(* IEC 61131-3 sources: plcassist-cli/packages/volt-lsp-iec/test-corpus/pro2193/Device/Plc Logic/Application/09 Misc/Library Manager/L_MC2P_MotionControlCam, 92 files *)

(* ---- L_MC2P_CONSTANTS.gvl ---- *)
VAR_GLOBAL
	GC_DWCHECKIDCOND : DWORD := 1000;
	GC_DWCHECKIDCHAR : DWORD := 2000;
	GC_DWCHECKIDDATAXYA : DWORD := 3000;
	GC_DWCHECKIDDATAXY : DWORD := 3500;
	GC_DWCHECKIDDATAYA : DWORD := 4000;
	GC_DWCHECKIDDATAY : DWORD := 4500;
	GC_DWCHECKIDCAMDATA : DWORD := 5000;
	GC_DWCHECKIDSCCAMTABLEID : DWORD := 6000;
	GC_DWCHECKIDCAMID : DWORD := 7000;
	GC_DWCHECKIDCAMREF : DWORD := 12000;
	GC_DWCHECKIDTAPPET : DWORD := 8000;
	GC_DWCHECKIDTAPPETDATA : DWORD := 9000;
	GC_DWCHECKIDTAPPETREF : DWORD := 10000;
	GC_DWCHECKIDTAPPETID : DWORD := 11000;
	GC_DWCHECKIDTAPPETPOS : DWORD := 11001;
	GC_DWCHECKIDTAPPETTIME : DWORD := 11002;
	GC_LRCORRECTCONDITIONPOSITION : LREAL := 1E-06;
	GC_UIBLOCKEDNUMOFCYCLES : UINT := 10;
END_VAR

(* ---- L_MC2P_EVENTS.gvl ---- *)
VAR_GLOBAL
	CMPID_EVT_NEWCAMFILESDOWNLOADED : UDINT := 16#2003;
	EVT_CMPLENZEIPCSYSTEMNEWCAMFILESDOWNLOADED : UDINT := 16#10001;
	EVTPARAMID_CMPLENZEIPCSYSTEMNEWCAMFILESDOWNLOADED : UDINT := 16#1;
	EVTVERSION_CMPLENZEIPCSYSTEMNEWCAMFILESDOWNLOADED : UDINT := 16#1;
END_VAR

(* ---- L_MC2P_INTERNALCONST.gvl ---- *)
VAR_GLOBAL
	MAGICLML : DWORD := 16#46444D4C;
	MAGICCRPT : DWORD := 16#54505243;
	MAGICORGA : DWORD := 16#4147524F;
	MAGICEND : DWORD := 16#444E454C;
	MAGICCD : WORD := 16#4443;
	MAGICTD : WORD := 16#4454;
	C_CAM_CRC_BUFFERSIZE : DWORD := 96;
	CRC32TABLE : ARRAY [0..255] OF DWORD := [16#0, 16#77073096, 16#EE0E612C, 16#990951BA, 16#76DC419, 16#706AF48F, 16#E963A535, 16#9E6495A3, 16#EDB8832, 16#79DCB8A4, 16#E0D5E91E, 16#97D2D988, 16#9B64C2B, 16#7EB17CBD, 16#E7B82D07, 16#90BF1D91, 16#1DB71064, 16#6AB020F2, 16#F3B97148, 16#84BE41DE, 16#1ADAD47D, 16#6DDDE4EB, 16#F4D4B551, 16#83D385C7, 16#136C9856, 16#646BA8C0, 16#FD62F97A, 16#8A65C9EC, 16#14015C4F, 16#63066CD9, 16#FA0F3D63, 16#8D080DF5, 16#3B6E20C8, 16#4C69105E, 16#D56041E4, 16#A2677172, 16#3C03E4D1, 16#4B04D447, 16#D20D85FD, 16#A50AB56B, 16#35B5A8FA, 16#42B2986C, 16#DBBBC9D6, 16#ACBCF940, 16#32D86CE3, 16#45DF5C75, 16#DCD60DCF, 16#ABD13D59, 16#26D930AC, 16#51DE003A, 16#C8D75180, 16#BFD06116, 16#21B4F4B5, 16#56B3C423, 16#CFBA9599, 16#B8BDA50F, 16#2802B89E, 16#5F058808, 16#C60CD9B2, 16#B10BE924, 16#2F6F7C87, 16#58684C11, 16#C1611DAB, 16#B6662D3D, 16#76DC4190, 16#1DB7106, 16#98D220BC, 16#EFD5102A, 16#71B18589, 16#6B6B51F, 16#9FBFE4A5, 16#E8B8D433, 16#7807C9A2, 16#F00F934, 16#9609A88E, 16#E10E9818, 16#7F6A0DBB, 16#86D3D2D, 16#91646C97, 16#E6635C01, 16#6B6B51F4, 16#1C6C6162, 16#856530D8, 16#F262004E, 16#6C0695ED, 16#1B01A57B, 16#8208F4C1, 16#F50FC457, 16#65B0D9C6, 16#12B7E950, 16#8BBEB8EA, 16#FCB9887C, 16#62DD1DDF, 16#15DA2D49, 16#8CD37CF3, 16#FBD44C65, 16#4DB26158, 16#3AB551CE, 16#A3BC0074, 16#D4BB30E2, 16#4ADFA541, 16#3DD895D7, 16#A4D1C46D, 16#D3D6F4FB, 16#4369E96A, 16#346ED9FC, 16#AD678846, 16#DA60B8D0, 16#44042D73, 16#33031DE5, 16#AA0A4C5F, 16#DD0D7CC9, 16#5005713C, 16#270241AA, 16#BE0B1010, 16#C90C2086, 16#5768B525, 16#206F85B3, 16#B966D409, 16#CE61E49F, 16#5EDEF90E, 16#29D9C998, 16#B0D09822, 16#C7D7A8B4, 16#59B33D17, 16#2EB40D81, 16#B7BD5C3B, 16#C0BA6CAD, 16#EDB88320, 16#9ABFB3B6, 16#3B6E20C, 16#74B1D29A, 16#EAD54739, 16#9DD277AF, 16#4DB2615, 16#73DC1683, 16#E3630B12, 16#94643B84, 16#D6D6A3E, 16#7A6A5AA8, 16#E40ECF0B, 16#9309FF9D, 16#A00AE27, 16#7D079EB1, 16#F00F9344, 16#8708A3D2, 16#1E01F268, 16#6906C2FE, 16#F762575D, 16#806567CB, 16#196C3671, 16#6E6B06E7, 16#FED41B76, 16#89D32BE0, 16#10DA7A5A, 16#67DD4ACC, 16#F9B9DF6F, 16#8EBEEFF9, 16#17B7BE43, 16#60B08ED5, 16#D6D6A3E8, 16#A1D1937E, 16#38D8C2C4, 16#4FDFF252, 16#D1BB67F1, 16#A6BC5767, 16#3FB506DD, 16#48B2364B, 16#D80D2BDA, 16#AF0A1B4C, 16#36034AF6, 16#41047A60, 16#DF60EFC3, 16#A867DF55, 16#316E8EEF, 16#4669BE79, 16#CB61B38C, 16#BC66831A, 16#256FD2A0, 16#5268E236, 16#CC0C7795, 16#BB0B4703, 16#220216B9, 16#5505262F, 16#C5BA3BBE, 16#B2BD0B28, 16#2BB45A92, 16#5CB36A04, 16#C2D7FFA7, 16#B5D0CF31, 16#2CD99E8B, 16#5BDEAE1D, 16#9B64C2B0, 16#EC63F226, 16#756AA39C, 16#26D930A, 16#9C0906A9, 16#EB0E363F, 16#72076785, 16#5005713, 16#95BF4A82, 16#E2B87A14, 16#7BB12BAE, 16#CB61B38, 16#92D28E9B, 16#E5D5BE0D, 16#7CDCEFB7, 16#BDBDF21, 16#86D3D2D4, 16#F1D4E242, 16#68DDB3F8, 16#1FDA836E, 16#81BE16CD, 16#F6B9265B, 16#6FB077E1, 16#18B74777, 16#88085AE6, 16#FF0F6A70, 16#66063BCA, 16#11010B5C, 16#8F659EFF, 16#F862AE69, 16#616BFFD3, 16#166CCF45, 16#A00AE278, 16#D70DD2EE, 16#4E048354, 16#3903B3C2, 16#A7672661, 16#D06016F7, 16#4969474D, 16#3E6E77DB, 16#AED16A4A, 16#D9D65ADC, 16#40DF0B66, 16#37D83BF0, 16#A9BCAE53, 16#DEBB9EC5, 16#47B2CF7F, 16#30B5FFE9, 16#BDBDF21C, 16#CABAC28A, 16#53B39330, 16#24B4A3A6, 16#BAD03605, 16#CDD70693, 16#54DE5729, 16#23D967BF, 16#B3667A2E, 16#C4614AB8, 16#5D681B02, 16#2A6F2B94, 16#B40BBE37, 16#C30C8EA1, 16#5A05DF1B, 16#2D02EF8D];
	C_TAPPETS_BUFFERSIZE : DWORD := 23;
END_VAR

(* ---- L_MC2P_IMOTIONDATA.itf ---- *)
INTERFACE L_MC2P_IMOTIONDATA
END_INTERFACE

(* ---- L_MC2P_ITAPPETDATA.itf ---- *)
INTERFACE L_MC2P_ITAPPETDATA
END_INTERFACE

(* ---- L_MC2P_SETVALUES.itf ---- *)
INTERFACE L_MC2P_SETVALUES
END_INTERFACE

METHOD GETVALUES : LREAL
VAR_INPUT
	ESOURCE : MC_Source;
END_VAR
END_METHOD

(* ---- L_MC2P_TAPPET_REF.itf ---- *)
INTERFACE L_MC2P_TAPPET_REF
END_INTERFACE

METHOD GETID : DWORD
END_METHOD

METHOD GETTAPPETDATA : POINTER TO L_MC2P_TappetData
END_METHOD

METHOD SETCAMDATAACTIVE
VAR_INPUT
	XCAMACITVE : BOOL;
END_VAR
END_METHOD

METHOD SETMASTERVALUES
VAR_INPUT
	LRMASTERPOS : LREAL;
END_VAR
END_METHOD

(* ---- MC_CAM_REF.itf ---- *)
INTERFACE MC_CAM_REF
END_INTERFACE

METHOD GETCAMDATA : POINTER TO L_MC2P_CamData
END_METHOD

METHOD GETID : DWORD
END_METHOD

METHOD SETCAMDATAACTIVE
VAR_INPUT
	XCAMACITVE : BOOL;
END_VAR
END_METHOD

METHOD SETMASTERVALUES
VAR_INPUT
	LRMASTERPOS : LREAL;
END_VAR
END_METHOD

(* ---- GETBOOLEANPROPERTY.fun ---- *)
FUNCTION GETBOOLEANPROPERTY : BOOL
VAR_INPUT
	STKEY : WSTRING;
END_VAR
END_FUNCTION

(* ---- GETCOMPANY.fun ---- *)
FUNCTION GETCOMPANY : WSTRING
END_FUNCTION

(* ---- GETNUMBERPROPERTY.fun ---- *)
FUNCTION GETNUMBERPROPERTY : DINT
VAR_INPUT
	STKEY : WSTRING;
END_VAR
END_FUNCTION

(* ---- GETTEXTPROPERTY.fun ---- *)
FUNCTION GETTEXTPROPERTY : WSTRING
VAR_INPUT
	STKEY : WSTRING;
END_VAR
END_FUNCTION

(* ---- GETTEXTPROPERTY2.fun ---- *)
FUNCTION GETTEXTPROPERTY2 : POINTER TO WSTRING
VAR_INPUT
	STKEY : WSTRING;
END_VAR
END_FUNCTION

(* ---- GETTITLE.fun ---- *)
FUNCTION GETTITLE : WSTRING
END_FUNCTION

(* ---- GETVERSION.fun ---- *)
FUNCTION GETVERSION : VERSION
END_FUNCTION

(* ---- GETVERSIONPROPERTY.fun ---- *)
FUNCTION GETVERSIONPROPERTY : VERSION
VAR_INPUT
	STKEY : WSTRING;
END_VAR
END_FUNCTION

(* ---- L_MC2P_CAMGETDATA.fun ---- *)
FUNCTION L_MC2P_CAMGETDATA : POINTER TO BYTE
VAR_INPUT
	ITFCAMDATA : L_MC2P_IMotionData;
	IDX : UDINT;
	ECAMTYPE : L_MC2P_CamType;
END_VAR
END_FUNCTION

(* ---- L_MC2P_CAMGETDATA2.fun ---- *)
FUNCTION L_MC2P_CAMGETDATA2 : BOOL
VAR_INPUT
	ITFCAMDATA : L_MC2P_IMotionData;
	IDX1 : UDINT;
	IDX2 : UDINT;
	ECAMTYPE : L_MC2P_CamType;
END_VAR
VAR_OUTPUT
	PSCDATA1 : POINTER TO BYTE;
	PSCDATA2 : POINTER TO BYTE;
END_VAR
END_FUNCTION

(* ---- L_MC2P_CAMGETXVALUE2.fun ---- *)
FUNCTION L_MC2P_CAMGETXVALUE2 : BOOL
VAR_INPUT
	ITFCAMDATA : L_MC2P_IMotionData;
	IDX1 : UDINT;
	IDX2 : UDINT;
	ECAMTYPE : L_MC2P_CamType;
	LRMASTEP : LREAL;
	LRXSTART : LREAL;
END_VAR
VAR_OUTPUT
	LRX1 : LREAL;
	LRX2 : LREAL;
END_VAR
END_FUNCTION

(* ---- L_MC2P_CAMGETYVALUE2.fun ---- *)
FUNCTION L_MC2P_CAMGETYVALUE2 : BOOL
VAR_INPUT
	ITFCAMDATA : L_MC2P_IMotionData;
	IDX1 : UDINT;
	IDX2 : UDINT;
	ECAMTYPE : L_MC2P_CamType;
END_VAR
VAR_OUTPUT
	LRY1 : LREAL;
	LRY2 : LREAL;
END_VAR
END_FUNCTION

(* ---- L_MC2P_CHECK_CAMREFEQ.fun ---- *)
FUNCTION L_MC2P_CHECK_CAMREFEQ : BOOL
VAR_INPUT
	CAMREFNEW : MC_CAM_REF;
	CAMREFOLD : MC_CAM_REF;
END_VAR
END_FUNCTION

(* ---- L_MC2P_CHECK_CAMTABLECHANGED.fun ---- *)
FUNCTION L_MC2P_CHECK_CAMTABLECHANGED : BOOL
VAR_INPUT
	SCCAMTABLENEW : MC_Cam_REF;
	SCCAMTABLEOLD : MC_Cam_REF;
	SCCAMINFOOLD : L_MC2P_CamInfo;
END_VAR
END_FUNCTION

(* ---- L_MC2P_CHECK_CAMTABLEVALID.fun ---- *)
FUNCTION L_MC2P_CHECK_CAMTABLEVALID : BOOL
VAR_INPUT
	CAMTABLE : MC_Cam_REF;
END_VAR
END_FUNCTION

(* ---- L_MC2P_CONVERTPOSTOMODULOPOS.fun ---- *)
FUNCTION L_MC2P_CONVERTPOSTOMODULOPOS : LREAL
VAR_INPUT
	LRPOS : LREAL;
	LRPERIOD : LREAL;
END_VAR
END_FUNCTION

(* ---- L_MC2P_CONVERTPOSTOMODULOPOSEXTENDED.fun ---- *)
FUNCTION L_MC2P_CONVERTPOSTOMODULOPOSEXTENDED : LREAL
VAR_INPUT
	LRPOS : LREAL;
	LRPERIOD : LREAL;
END_VAR
END_FUNCTION

(* ---- L_MC2P_HLPMODULO.fun ---- *)
FUNCTION L_MC2P_HLPMODULO : LREAL
VAR_INPUT
	LRINPUT : LREAL;
	LRLENGHT : LREAL;
END_VAR
END_FUNCTION

(* ---- L_MC2P_HLPMODULOADD.fun ---- *)
FUNCTION L_MC2P_HLPMODULOADD : LREAL
VAR_INPUT
	LRINPUT : LREAL;
	LROFFSET : LREAL;
	LRLENGHT : LREAL;
END_VAR
END_FUNCTION

(* ---- L_MC2P_HLPMODULODIFF.fun ---- *)
FUNCTION L_MC2P_HLPMODULODIFF : LREAL
VAR_INPUT
	LRDIFF : LREAL;
	LRLEN : LREAL;
END_VAR
END_FUNCTION

(* ---- L_MC2P_HLPMODULOZERO.fun ---- *)
FUNCTION L_MC2P_HLPMODULOZERO : BOOL
VAR_INPUT
	LRDIFF : LREAL;
	LRLEN : LREAL;
END_VAR
END_FUNCTION

(* ---- CRYPTING.fb ---- *)
FUNCTION_BLOCK CRYPTING
END_FUNCTION_BLOCK

METHOD DECRYPTMODE1
VAR_INPUT
	NUM_CYCLES : WORD;
	V : POINTER TO ARRAY [0..1] OF UDINT;
	K : ARRAY [0..3] OF UDINT;
END_VAR
END_METHOD

METHOD DECRYPTMODE64
VAR_INPUT
	NUM_CYCLES : WORD;
	V : POINTER TO ARRAY [0..1] OF ULINT;
	K : ARRAY [0..3] OF ULINT;
END_VAR
END_METHOD

METHOD ENCRYPTMODE1
VAR_INPUT
	NUM_CYCLES : WORD;
	V : POINTER TO ARRAY [0..1] OF UDINT;
	K : ARRAY [0..3] OF UDINT;
END_VAR
END_METHOD

METHOD ENCRYPTMODE64
VAR_INPUT
	NUM_CYCLES : WORD;
	V : POINTER TO ARRAY [0..1] OF ULINT;
	K : ARRAY [0..3] OF ULINT;
END_VAR
END_METHOD

METHOD GETLINTFROMCHAR : ULINT
VAR_INPUT
	ABDATA : ARRAY [0..3] OF BYTE;
END_VAR
END_METHOD

METHOD SETKEY : ARRAY [0..3] OF ULINT
VAR_INPUT
	SSTRING : STRING(16);
END_VAR
END_METHOD

(* ---- GLOBALTEXTLIST.fb ---- *)
FUNCTION_BLOCK GLOBALTEXTLIST
VAR
	M_TEXTLISTFILE : STRING(255);
	_STNAMESPACE : STRING;
END_VAR
END_FUNCTION_BLOCK

(* ---- IMAGEPOOL.fb ---- *)
FUNCTION_BLOCK IMAGEPOOL
VAR
	M_STNAMESPACE : STRING(80);
	M_STHELPVARID : STRING;
	M_STHELPVARPATH : STRING(255);
	M_STHELP : STRING;
	M_REGISTERIMAGES : BOOL := TRUE;
END_VAR
END_FUNCTION_BLOCK

METHOD FB_INIT : BOOL
VAR_INPUT
	BINITRETAINS : BOOL;
	BINCOPYCODE : BOOL;
END_VAR
END_METHOD

METHOD FB_REINIT : BOOL
END_METHOD

METHOD FB_EXIT : BOOL
VAR_INPUT
	BINCOPYCODE : BOOL;
END_VAR
END_METHOD

(* ---- L_MC2P_AXISCONVERTERBASE.fb ---- *)
FUNCTION_BLOCK L_MC2P_AXISCONVERTERBASE EXTENDS L_MC2P_CamAxisConverter
VAR_INPUT
	XENABLE : BOOL;
	LRCYCMASTERPOS : LREAL;
	LRCYCMASTERVEL : LREAL;
	LRCYCMASTERACC : LREAL;
	LRCYCLELENGTHMASTER : LREAL := 360;
	IMASTERMOVEMENTTYPE : INT := 0;
	LRCYCLELENGTHSLAVE : LREAL := 360;
	ISLAVEMOVEMENTTYPE : INT := 0;
	LRSETOFFSET : LREAL;
	LRSETSCALING : LREAL := 1;
	ESCALINGMODE : L_MC2P_ScalingMode := L_MC2P_ScalingMode.absolute;
END_VAR
VAR_OUTPUT
	XERROR : BOOL;
	EERRORID : L_IE1P_Error;
	XBUSY : BOOL;
	LRSETSLAVEPOSOUT : LREAL;
	LRSETSLAVEVELOUT : LREAL;
	LRSETSLAVEACCOUT : LREAL;
END_VAR
VAR
	XERROR_OLD : BOOL;
	EERRORID_OLD : L_IE1P_Error;
	XENABLE_OLD : BOOL;
	LRCYCMASTERPOS_OLD : LREAL;
	ESTATE : L_MC2P_States := L_MC2P_States.INIT;
	XSTATEENTRY : BOOL;
	BYCONVERTERMODE : BYTE;
	SCSETSLAVEOUT : L_MC2P_AxisProfile;
END_VAR
END_FUNCTION_BLOCK

METHOD CALL_CONVERTLINEARTOLINEAR
END_METHOD

METHOD CALL_CONVERTLINEARTOMODULO
END_METHOD

METHOD CALL_CONVERTMODULOTOLINEAR
END_METHOD

METHOD CALL_CONVERTMODULOTOMODULO
END_METHOD

METHOD CALL_ERRORHANDLER
END_METHOD

METHOD CALL_FBMETHODS
END_METHOD

METHOD CALL_OUTPUT
END_METHOD

METHOD CALL_RESETCOMMANDS
END_METHOD

METHOD CALL_RESETOUTPUT
END_METHOD

METHOD CALL_STATEMASHINE
END_METHOD

METHOD CALL_S000_CYCLIC
END_METHOD

METHOD CALL_S001_INIT
END_METHOD

METHOD CALL_S010_READY
END_METHOD

METHOD CALL_S200_SYNCHRON
END_METHOD

METHOD CALL_S998_ERROR
END_METHOD

(* ---- L_MC2P_BOUNDSCAM.fb ---- *)
FUNCTION_BLOCK L_MC2P_BOUNDSCAM EXTENDS L_MC2P_TemplateSlaveAxis
VAR_INPUT
	XEXECUTE : BOOL;
	ITFCAMTABLE : MC_CAM_REF;
	LRMAVEL : LREAL;
	LRMAACC : LREAL;
	UDINUMOFPOINTS : UDINT;
	UDIPOINTSPERCYCLE : UDINT;
END_VAR
VAR_OUTPUT
	XDONE : BOOL;
	XBUSY : BOOL;
	XERROR : BOOL;
	EERRORID : L_IE1P_Error;
	LRPOSMAX : LREAL;
	LRPOSMIN : LREAL;
	LRVELMAX : LREAL;
	LRVELMIN : LREAL;
	LRACCDECMAX : LREAL;
	LRACCDECMIN : LREAL;
END_VAR
VAR
	L_MC2P_CAMBASIC1 : L_MC2P_CamBasic;
	SCVIRTUALSLAVE : L_MC2P_AxisProfile;
	I : UDINT;
	LRMASTEP : LREAL;
	LRMAPOS : LREAL;
	XBREAK : BOOL;
	XEXECUTEOLD : BOOL;
	XRESETOUTPUT : BOOL;
	SCVIRTUALMASTER : L_MC2P_AxisProfile;
	LRMAVEL_INT : LREAL;
	LRMAACC_INT : LREAL;
	UDINUMOFPOINTS_INT : UDINT := 2;
	UDIPOINTSPERCYCLE_INT : UDINT;
	PCAMDATA_INT : POINTER TO L_MC2P_CamData;
	SCCAMINFO : L_MC2P_CamInfo;
	LRPOSMAX_INT : LREAL;
	LRPOSMIN_INT : LREAL;
	LRVELMAX_INT : LREAL;
	LRVELMIN_INT : LREAL;
	LRACCDECMAX_INT : LREAL;
	LRACCDECMIN_INT : LREAL;
END_VAR
END_FUNCTION_BLOCK

METHOD READINPUTS
END_METHOD

METHOD RESET_MINMAXVALUES
END_METHOD

METHOD RESET_OUTPUTS
END_METHOD

METHOD RESET_OUTPUTSBYERROR
END_METHOD

METHOD SET_MINMAXVALUES
END_METHOD

(* ---- L_MC2P_CAMAXISCONVERTER.fb ---- *)
FUNCTION_BLOCK L_MC2P_CAMAXISCONVERTER
VAR
	_XERROR : BOOL;
	LRSLAVEPERIOD_INT : LREAL := 0;
	LRSETSLAVEPOSOUTSCALED : LREAL := 0;
	DWACTSLAVEPOS_INT : DWORD := 0;
	LRSETSLAVEPOSOUT_INT : LREAL := 0;
	LRSLAVEOFFSET_INT : LREAL := 0;
	LRSLAVEOFFSET_REL : LREAL := 0;
	LRYOFFSET_INT : LREAL := 0;
	LRSETYPOS_INT : LREAL := 0;
	LRSETYPOS_SCALED : LREAL := 0;
	LRSETYSCALING_INT : LREAL := 1;
	ALRMEM : ARRAY [1..7] OF LREAL;
	XMODULOMODE : BOOL;
	LRXPERIOD_NEXT : LREAL;
	LRSTARTXAXIS_NEXT : LREAL := 0;
	LRSETXPOSOUT_MODULO : LREAL := 0;
	LRSETXPOSOUT_MODULO_OLD : LREAL := 0;
	LRSETXPOSOUT_INT : LREAL := 0;
	LRXPERIOD_INT : LREAL := 0;
	LRSTARTXAXIS_INT : LREAL := 0;
	LRSETXSCALING_INT : LREAL := 1;
	LROFFSET_INT : LREAL := 0;
	LROFFSET_REL : LREAL := 0;
	LRONECYCLEXOFFSET_INT : LREAL := 0;
	XLOADSTARTXPOS : BOOL;
	LRLOADSTARTXPOS : LREAL;
	XCHECKMASTERPOSBYLOAD : BOOL;
	LRCYCSETMASTERPOSBYLOAD : LREAL;
	LRSETXPOSBYLOAD : LREAL;
	XOVERRUNMASTERPOS : BOOL := FALSE;
	XOVERRUNMASTERNEG : BOOL := FALSE;
	LWREMAINDER_ADD : LWORD := 0;
	LWREMAINDER_INT : LWORD := 0;
	LRREMAINDER_INT : LREAL := 0;
	LRCYCSETMASTERPOS_VIRTUAL : LREAL := 0;
	LRMASTERPERIOD_VIRTUAL : LREAL := 0;
	IPERIODFACTOR : INT := 0;
	IPERIODCTN : INT := 0;
	LRCYCSETMASTERVEL_INT : LREAL;
	LRCYCSETMASTERPOS_INT : LREAL;
	LRMASTERPERIOD_INT : LREAL := 0;
	LRCYCSETMASTERPOS_SCALED : LREAL := 0;
	LRMASTERPERIOD_SCALED : LREAL := 0;
	XEOP_INIT : BOOL := TRUE;
	IEOP_CYCLECNTR : INT := 0;
	IEOP_CYCLECNTR2 : INT := 0;
	LWEOP_TCHECKSUM : LWORD;
	XEOP_ENDOFPERIODPOSITIVE : BOOL;
	XEOP_ENDOFPERIODNEGATIVE : BOOL;
	WEOP_STEPPER : WORD := 0;
	LREOP_CYCSETMASTERPOS_OLD : LREAL;
	LREOP_SETXPOSOUT_MODULO_OLD : LREAL;
	LREOP_XPERIOD : LREAL;
	LREOP_XPERIOD_OLD : LREAL;
	XEOP_ENDOFPROFPOSITIVE : BOOL;
	XEOP_ENDOFPROFNEGATIVE : BOOL;
	LREOP_SETXDELTAPOS : LREAL;
	LREOP_SETXDELTA2POS : LREAL;
	LREOP_SETXDELTA3POS : LREAL;
	LREOP_SETXDELTAPOS_OLD : LREAL;
	LREOP_SETXDELTA2POS_OLD : LREAL;
	LREOP_SETXSCALING_OLD : LREAL;
	LREOP_OFFSET_OLD : LREAL;
	ALREOP_MEM : ARRAY [1..7] OF LREAL;
	XEOP_RAMPOFFSETMODE : BOOL;
	XEOP_RAMPSCALINGMODE : BOOL;
	XOUTOFCAMPOSITIVE_INT : BOOL;
	XOUTOFCAMNEGATIVE_INT : BOOL;
	LRTEMP : LREAL;
	LRENDOFPROFILEFACTOR_INT : LREAL := 1;
	LRCYCSETMASTERPOSATSCLING0 : LREAL;
	LRSETXPOSOUTATSCLING0 : LREAL;
	LRSETXSCALINGATSCLING0 : LREAL;
	LRDWUPPERLIMIT : LREAL := 16#FFFFFFFF;
	DWDWUPPERLIMIT : DWORD := 16#FFFFFFFF;
	LRLWUPPERLIMIT : LREAL := 16#7FFFFFFFFFFFFFFF;
	LWENDOFPROFILECHECKSUM : LWORD;
END_VAR
END_FUNCTION_BLOCK

METHOD CALC_LRSETSLAVEPOSOUT : LREAL
VAR_IN_OUT
	LRSETYPOS : LREAL;
END_VAR
END_METHOD

METHOD CALC_LRSETXLINPOSOUT : LREAL
VAR_IN_OUT
	LRCYCSETMASTERPOS : LREAL;
	LRCYCSETMASTERVEL : LREAL;
	LRCYCSETMASTERACC : LREAL;
END_VAR
END_METHOD

METHOD CALC_LRSETXPOSOUT : LREAL
VAR_IN_OUT
	LRCYCSETMASTERPOS : LREAL;
	LRCYCSETMASTERVEL : LREAL;
	LRCYCSETMASTERACC : LREAL;
END_VAR
END_METHOD

METHOD CALC_LRSETXPOSOUTEXTENDED : LREAL
VAR_INPUT
	LRENDOFPROFILEWINDOW : LREAL;
END_VAR
VAR_OUTPUT
	LRSETXPOSOUT : LREAL;
	XENDOFPROFPOSITIVE : BOOL;
	XENDOFPROFNEGATIVE : BOOL;
	XEXTRAPOLATECAM : BOOL;
	XCYCLEZERO : BOOL;
	XOUTOFCAMPOSITIVE : BOOL;
	XOUTOFCAMNEGATIVE : BOOL;
END_VAR
VAR_IN_OUT
	LRCYCSETMASTERPOS : LREAL;
	LRCYCSETMASTERPOS_OLD : LREAL;
	LRCYCSETMASTERVEL : LREAL;
	LRCYCSETMASTERACC : LREAL;
END_VAR
END_METHOD

METHOD CALL_RESET
END_METHOD

METHOD SET_LRENDOFPROFILEFACTOR : BOOL
VAR_INPUT
	LRIN : LREAL;
END_VAR
END_METHOD

METHOD CALC_DWADDMODULO : DWORD
VAR_INPUT
	LRSETXPOS : LREAL;
	LRSETYPOS : LREAL;
	LRPERIOD : LREAL;
END_VAR
END_METHOD

METHOD CALC_DWSUBMODULO : DWORD
VAR_INPUT
	LRSETYPOS : LREAL;
	LRSETXPOS : LREAL;
	LRPERIOD : LREAL;
END_VAR
END_METHOD

METHOD CALC_LRADDMODULO : LREAL
VAR_INPUT
	LRSETXPOS : LREAL;
	LRSETYPOS : LREAL;
	LRPERIOD : LREAL;
END_VAR
END_METHOD

METHOD CALC_LRSUBMODULO : LREAL
VAR_INPUT
	LRSETXPOS : LREAL;
	LRSETYPOS : LREAL;
	LRPERIOD : LREAL;
END_VAR
END_METHOD

METHOD CALL_CHECKLOADXPOSAFTERCONVERTER
END_METHOD

METHOD CALL_CHECKMODULOOVERRUN
VAR_IN_OUT
	LRSETPOS : LREAL;
	LRSETVEL : LREAL;
	LRPERIOD : LREAL;
	XOVERRUNPOS : BOOL;
	XOVERRUNNEG : BOOL;
	ALRMEM : ARRAY [1..7] OF LREAL;
END_VAR
END_METHOD

METHOD CALL_DWCONVERTLREALTODWORD : DWORD
VAR_INPUT
	LRIN : LREAL;
	LRPERIOD : LREAL;
END_VAR
END_METHOD

METHOD CALL_DWCONVERTLREALTOLWORD : LWORD
VAR_INPUT
	LRIN : LREAL;
	LRPERIOD : LREAL;
END_VAR
END_METHOD

METHOD CALL_LRCONVERTDWORDTOLREAL : LREAL
VAR_INPUT
	DWIN : DWORD;
	LRPERIOD : LREAL;
END_VAR
END_METHOD

METHOD CALL_LRCONVERTLREALTOMODULO : LREAL
VAR_INPUT
	LRIN : LREAL;
	LRPERIOD : LREAL;
END_VAR
END_METHOD

METHOD CALL_LRCONVERTLWORDTOLREAL : LREAL
VAR_INPUT
	LWIN : LWORD;
	LRPERIOD : LREAL;
END_VAR
END_METHOD

METHOD CALC_MASTERVIRTUALPERIOD
END_METHOD

METHOD CALL_CHECKMODULOMODE
END_METHOD

METHOD CALL_CHECKZERROPOS
VAR_INPUT
	LRCYCSETMASTERPOS : LREAL;
END_VAR
END_METHOD

METHOD CHECK_XENDOFPROFILE : BOOL
VAR_INPUT
	LRSETXPOS : LREAL;
	LRSETXDELTAPOS : LREAL;
	LRSETXDELTA2POS : LREAL;
	LRSETXDELTA3POS : LREAL;
	LRXSTART : LREAL;
	LRXEND : LREAL;
	LRXPERIOD : LREAL;
END_VAR
VAR_OUTPUT
	LRSETNEXTXPOSOUT : LREAL;
	XPOSITIVE : BOOL;
	XNEGATIVE : BOOL;
END_VAR
END_METHOD

METHOD CALL_XMASTERVALID : BOOL
END_METHOD

METHOD GET_LRSLAVEOFFSETREL : LREAL
END_METHOD

METHOD GET_LRXOFFSETREL : LREAL
END_METHOD

METHOD LOAD_STARTXPOS
VAR_IN_OUT
	LRLOADXPOS : LREAL;
	LRCYCSETMASTERPOS : LREAL;
END_VAR
END_METHOD

METHOD SET_ACTAXISLIMIT
VAR_IN_OUT
	LRSTARTXAXIS : LREAL := 0;
	LRENDXAXIS : LREAL := 0;
END_VAR
END_METHOD

METHOD SET_EOPXOFFSETMODE
VAR_INPUT
	XRAMPOFFSETMODE : BOOL;
END_VAR
END_METHOD

METHOD SET_EOPXSCALINGMODE
VAR_INPUT
	XRAMPSCALINGMODE : BOOL;
END_VAR
END_METHOD

METHOD SET_NEWXPERIOD
VAR_IN_OUT
	LRSETXPOSOUT : LREAL;
	LRSETXPERIOD : LREAL;
	LRCYCSETMASTERPOS : LREAL;
END_VAR
END_METHOD

METHOD SET_NEXTAXISLIMIT
VAR_IN_OUT
	LRSTARTXAXIS : LREAL := 0;
	LRENDXAXIS : LREAL := 0;
END_VAR
END_METHOD

METHOD SET_ONECYCLEOFFSET
VAR_INPUT
	LRXOFFSET : LREAL;
END_VAR
END_METHOD

METHOD SET_XAXISLIMIT
VAR_INPUT
	LRSTARTXAXIS : LREAL;
	LRENDXAXIS : LREAL;
	LRSETSCALING : LREAL;
END_VAR
END_METHOD

METHOD SET_XOFFSET
VAR_INPUT
	LRSETOFFSET : LREAL;
END_VAR
END_METHOD

METHOD SET_XPERIOD
VAR_IN_OUT
	LRXPERIOD : LREAL;
	LRSETSCALING : LREAL;
END_VAR
END_METHOD

METHOD SET_XPOSTOMASTERPOS : DWORD
VAR_IN_OUT
	LRCYCSETMASTERPOS : LREAL;
END_VAR
END_METHOD

METHOD SET_XSCALING
VAR_INPUT
	LRSETSCALING : LREAL := 1;
	WSCALINGMODE : WORD := 0;
	LRCYCSETMASTERPOS : LREAL;
	LRCYCSETMASTERPOS_OLD : LREAL;
END_VAR
END_METHOD

METHOD SET_LRMASTERPERIOD
VAR_INPUT
	LRSETMASTERPERIOD : LREAL;
END_VAR
END_METHOD

METHOD LOAD_SALVEPOS
VAR_INPUT
	LRLOADSLAVEPOS : LREAL;
	LRSETYPOS : LREAL;
	LRSETYSCALING : LREAL;
END_VAR
END_METHOD

METHOD SET_SLAVEPOSTOYPOS : DWORD
VAR_INPUT
	LRSETYSCALING : LREAL;
END_VAR
END_METHOD

METHOD SET_YSCALING
VAR_INPUT
	LRSETSCALING : LREAL := 1;
	WSCALINGMODE : WORD := 0;
	LRSETSLAVEPOSOUT : LREAL;
	LRSETYPOS_OLD : LREAL;
END_VAR
END_METHOD

METHOD SET_LRCAMPOSDIFF
VAR_INPUT
	LRCAMPOSDIFF : LREAL;
END_VAR
END_METHOD

METHOD SET_LRCAMSWITCHREL
VAR_INPUT
	XDIRECTIONPOS : BOOL;
	LRYSCALINGEND : LREAL;
	LRYSCALINGSTART : LREAL;
	LRCAMYEND : LREAL;
	LRCAMYSTART : LREAL;
END_VAR
END_METHOD

METHOD SET_LRSLAVEOFFSET
VAR_INPUT
	LRSETOFFSET : LREAL;
END_VAR
END_METHOD

METHOD SET_LRSLAVEPERIOD
VAR_INPUT
	LRSETSLAVEPERIOD : LREAL;
END_VAR
END_METHOD

METHOD SET_LRYOFFSET
VAR_INPUT
	LRSETOFFSET : LREAL;
END_VAR
END_METHOD

(* ---- L_MC2P_CAMBASIC.fb ---- *)
FUNCTION_BLOCK L_MC2P_CAMBASIC
VAR
	LRENDVEL : LREAL;
	LRSTARTVEL : LREAL;
	LRENDACC : LREAL;
	LRSTARTACC : LREAL;
	LRMASTEP : LREAL;
	UDISEG : UDINT;
	UDISEGOLD : UDINT;
	UDISEGADD2 : UDINT;
	UDISEGSUB1 : UDINT;
	UDILEFTBORDER : UDINT;
	UDIRIGHTBORDER : UDINT;
	XFOUNDSEG : BOOL;
	SCCHAR : ARRAY [0..1] OF L_MC2P_Characteristics;
	WDEBUG : WORD;
	XRESTARTSERCH : BOOL;
	LRMAPOSOLD : LREAL;
	PCAMDATAOLD : POINTER TO BYTE;
	PDATAOLD : POINTER TO BYTE;
	ECAMTYPEOLD : DWORD;
	UDINUMOFELEMENTSOLD : DWORD;
	LRXSTARTPOSOLD : LREAL;
	LRXENDPOSOLD : LREAL;
	WSLAVESTATEOLDCYCLE : WORD;
	WSLAVESTATEOLDCAM : WORD;
	SCOUTPUTSLAVEOLDCYCLE : L_MC2P_AxisProfile;
	XNEWCAMDETECTED : BOOL;
	ACTUALSEGMENT : UDINT;
	FOUNDSEG : BOOL;
END_VAR
END_FUNCTION_BLOCK

METHOD CALCULATECAMPROFILE
VAR_INPUT
	PCAMDATA : POINTER TO L_MC2P_CamData;
	SCINPUTMASTER : L_MC2P_AxisProfile;
	XPERIODIC : BOOL;
	XEXTRAPOLATECAM : BOOL;
END_VAR
VAR_OUTPUT
	SCOUTPUTSLAVE : L_MC2P_AxisProfile;
	XERROR : BOOL;
	EERRORID : L_IE1P_Error;
END_VAR
END_METHOD

METHOD CALCULATECAMPROFILEINT
VAR_INPUT
	PCAMDATA : POINTER TO L_MC2P_CamData;
	SCINPUTMASTER : L_MC2P_AxisProfile;
	XPERIODIC : BOOL;
END_VAR
VAR_OUTPUT
	SCOUTPUTSLAVE : L_MC2P_AxisProfile;
	XERROR : BOOL;
	EERRORID : L_IE1P_Error;
END_VAR
END_METHOD

METHOD CAMGENERATORCOND
VAR_INPUT
	ITFCAMDATA : L_MC2P_IMotionData;
	LRINPUTMASTERVEL : LREAL;
	PSCCHAR : POINTER TO L_MC2P_Characteristics;
END_VAR
VAR_OUTPUT
	XERROR : BOOL;
	EERRORID : L_IE1P_Error;
END_VAR
END_METHOD

METHOD CAMPROFILERCHARCALC
VAR_INPUT
	PSCCHAR : POINTER TO L_MC2P_Characteristics;
	LRPOS : LREAL;
	UDISEGCHAR : UDINT;
	LRINPUTMASTERVEL : LREAL;
	LRINPUTMASTERACC : LREAL;
END_VAR
VAR_OUTPUT
	SCOUTPUTSLAVE : L_MC2P_AxisProfile;
END_VAR
END_METHOD

METHOD CAMPROFILERCHARSEARCH
VAR_INPUT
	PSCCHAR : POINTER TO L_MC2P_Characteristics;
	LRINPUTMASTERPOS : LREAL;
	ECAMTYPE : L_MC2P_CamType;
END_VAR
VAR_OUTPUT
	LRPOS : LREAL;
	UDISEGCHAR : UDINT;
END_VAR
END_METHOD

METHOD CAMPROFILERDATAEQUIY
VAR_INPUT
	PCAMDATA : POINTER TO L_MC2P_CamData;
	LRINPUTMASTERPOS : LREAL;
	LRINPUTMASTERVEL : LREAL;
	LRINPUTMASTERACC : LREAL;
	XPERIODIC : BOOL;
END_VAR
VAR_OUTPUT
	SCOUTPUTSLAVE : L_MC2P_AxisProfile;
	XERROR : BOOL;
	EERRORID : L_IE1P_Error;
END_VAR
END_METHOD

METHOD CAMPROFILERDATAEQUIYA
VAR_INPUT
	PCAMDATA : POINTER TO L_MC2P_CamData;
	LRINPUTMASTERPOS : LREAL;
	LRINPUTMASTERVEL : LREAL;
	LRINPUTMASTERACC : LREAL;
	XPERIODIC : BOOL;
END_VAR
VAR_OUTPUT
	SCOUTPUTSLAVE : L_MC2P_AxisProfile;
	XERROR : BOOL;
	EERRORID : L_IE1P_Error;
END_VAR
END_METHOD

METHOD CAMPROFILERDATANONEQUIXY
VAR_INPUT
	PCAMDATA : POINTER TO L_MC2P_CamData;
	LRINPUTMASTERPOS : LREAL;
	LRINPUTMASTERVEL : LREAL;
	LRINPUTMASTERACC : LREAL;
	XPERIODIC : BOOL;
END_VAR
VAR_OUTPUT
	SCOUTPUTSLAVE : L_MC2P_AxisProfile;
	XERROR : BOOL;
	EERRORID : L_IE1P_Error;
END_VAR
END_METHOD

METHOD CAMPROFILERDATANONEQUIXYA
VAR_INPUT
	PCAMDATA : POINTER TO L_MC2P_CamData;
	LRINPUTMASTERPOS : LREAL;
	LRINPUTMASTERVEL : LREAL;
	LRINPUTMASTERACC : LREAL;
	XPERIODIC : BOOL;
END_VAR
VAR_OUTPUT
	SCOUTPUTSLAVE : L_MC2P_AxisProfile;
	XERROR : BOOL;
	EERRORID : L_IE1P_Error;
END_VAR
END_METHOD

METHOD GETSTARTENDVALUES
VAR_INPUT
	PCAMDATA : POINTER TO L_MC2P_CamData;
END_VAR
VAR_OUTPUT
	LRSTARTSLAVE : LREAL;
	LRENDSLAVE : LREAL;
END_VAR
END_METHOD

METHOD RESETSEGMENT
END_METHOD

METHOD SEARCHSEGMENT
VAR_INPUT
	PCAMDATA : POINTER TO L_MC2P_CamData;
	LRINPUTMASTERPOS : LREAL;
	LRINPUTMASTERVEL : LREAL;
	XPERIODIC : BOOL;
END_VAR
VAR_OUTPUT
	XERROR : BOOL;
	EERRORID : L_IE1P_Error;
END_VAR
END_METHOD

METHOD FB_INIT : BOOL
VAR_INPUT
	BINITRETAINS : BOOL;
	BINCOPYCODE : BOOL;
END_VAR
END_METHOD

METHOD GETEXTREMVALUES_POLY5
VAR_INPUT
	PSCCHARCLUTCH : POINTER TO L_MC2P_Characteristics;
END_VAR
VAR_OUTPUT
	LRFSMAX1 : LREAL;
	LRFSMAX2 : LREAL;
	LRFSMAX3 : LREAL;
END_VAR
END_METHOD

METHOD GEN_BB_POLY5
VAR_INPUT
	PSCCONDLEFT : POINTER TO L_MC2P_XYVA;
	PSCCONDRIGHT : POINTER TO L_MC2P_XYVA;
	PSCCHAR : POINTER TO L_MC2P_Characteristics;
END_VAR
END_METHOD

METHOD GEN_BB_POLY7
VAR_INPUT
	PSCCONDLEFT : POINTER TO L_MC2P_XYVA;
	PSCCONDRIGHT : POINTER TO L_MC2P_XYVA;
	PSCCHAR : POINTER TO L_MC2P_Characteristics;
END_VAR
END_METHOD

METHOD GEN_GG_GERADE
VAR_INPUT
	PSCCONDLEFT : POINTER TO L_MC2P_XYVA;
	PSCCONDRIGHT : POINTER TO L_MC2P_XYVA;
	PSCCHAR : POINTER TO L_MC2P_Characteristics;
END_VAR
END_METHOD

METHOD GEN_GG_MODSIN
VAR_INPUT
	PSCCONDLEFT : POINTER TO L_MC2P_XYVA;
	PSCCONDRIGHT : POINTER TO L_MC2P_XYVA;
	PSCCHAR : POINTER TO L_MC2P_Characteristics;
END_VAR
END_METHOD

METHOD GEN_GG_POLY3
VAR_INPUT
	PSCCONDLEFT : POINTER TO L_MC2P_XYVA;
	PSCCONDRIGHT : POINTER TO L_MC2P_XYVA;
	PSCCHAR : POINTER TO L_MC2P_Characteristics;
END_VAR
END_METHOD

METHOD GEN_GR_POLY2
VAR_INPUT
	PSCCONDLEFT : POINTER TO L_MC2P_XYVA;
	PSCCONDRIGHT : POINTER TO L_MC2P_XYVA;
	PSCCHAR : POINTER TO L_MC2P_Characteristics;
END_VAR
END_METHOD

METHOD GEN_GU_HARMKOMB
VAR_INPUT
	PSCCONDLEFT : POINTER TO L_MC2P_XYVA;
	PSCCONDRIGHT : POINTER TO L_MC2P_XYVA;
	PSCCHAR : POINTER TO L_MC2P_Characteristics;
END_VAR
END_METHOD

METHOD GEN_RG_POLY2
VAR_INPUT
	PSCCONDLEFT : POINTER TO L_MC2P_XYVA;
	PSCCONDRIGHT : POINTER TO L_MC2P_XYVA;
	PSCCHAR : POINTER TO L_MC2P_Characteristics;
END_VAR
END_METHOD

METHOD GEN_RR_BESCHLTRAPEZ
VAR_INPUT
	PSCCONDLEFT : POINTER TO L_MC2P_XYVA;
	PSCCONDRIGHT : POINTER TO L_MC2P_XYVA;
	PSCCHAR : POINTER TO L_MC2P_Characteristics;
END_VAR
END_METHOD

METHOD GEN_RR_GENSIN
VAR_INPUT
	PSCCONDLEFT : POINTER TO L_MC2P_XYVA;
	PSCCONDRIGHT : POINTER TO L_MC2P_XYVA;
	PSCCHAR : POINTER TO L_MC2P_Characteristics;
END_VAR
END_METHOD

METHOD GEN_RR_MODBESCHLTRAPEZ
VAR_INPUT
	PSCCONDLEFT : POINTER TO L_MC2P_XYVA;
	PSCCONDRIGHT : POINTER TO L_MC2P_XYVA;
	PSCCHAR : POINTER TO L_MC2P_Characteristics;
END_VAR
END_METHOD

METHOD GEN_RR_QUADPARABEL
VAR_INPUT
	PSCCONDLEFT : POINTER TO L_MC2P_XYVA;
	PSCCONDRIGHT : POINTER TO L_MC2P_XYVA;
	PSCCHAR : POINTER TO L_MC2P_Characteristics;
END_VAR
END_METHOD

METHOD GEN_RR_SIN
VAR_INPUT
	PSCCONDLEFT : POINTER TO L_MC2P_XYVA;
	PSCCONDRIGHT : POINTER TO L_MC2P_XYVA;
	PSCCHAR : POINTER TO L_MC2P_Characteristics;
END_VAR
END_METHOD

METHOD GEN_RU_MODBESCHLTRAPEZ
VAR_INPUT
	PSCCONDLEFT : POINTER TO L_MC2P_XYVA;
	PSCCONDRIGHT : POINTER TO L_MC2P_XYVA;
	PSCCHAR : POINTER TO L_MC2P_Characteristics;
END_VAR
END_METHOD

METHOD GEN_UG_HARMKOMB
VAR_INPUT
	PSCCONDLEFT : POINTER TO L_MC2P_XYVA;
	PSCCONDRIGHT : POINTER TO L_MC2P_XYVA;
	PSCCHAR : POINTER TO L_MC2P_Characteristics;
END_VAR
END_METHOD

METHOD GEN_UR_MODBESCHLTRAPEZ
VAR_INPUT
	PSCCONDLEFT : POINTER TO L_MC2P_XYVA;
	PSCCONDRIGHT : POINTER TO L_MC2P_XYVA;
	PSCCHAR : POINTER TO L_MC2P_Characteristics;
END_VAR
END_METHOD

METHOD GEN_UU_SINGERKOMB : ARRAY [0..1] OF L_MC2P_Characteristics
VAR_INPUT
	PSCCONDLEFT : POINTER TO L_MC2P_XYVA;
	PSCCONDRIGHT : POINTER TO L_MC2P_XYVA;
	PSCCHAR : POINTER TO L_MC2P_Characteristics;
END_VAR
END_METHOD

METHOD PROF_BB_POLY5
VAR_INPUT
	PSCCHAR : POINTER TO L_MC2P_Characteristics;
	LRPOS : LREAL;
	PSCNORMSLAVE : POINTER TO L_MC2P_AxisProfile;
END_VAR
END_METHOD

METHOD PROF_BB_POLY7
VAR_INPUT
	PSCCHAR : POINTER TO L_MC2P_Characteristics;
	LRPOS : LREAL;
	PSCNORMSLAVE : POINTER TO L_MC2P_AxisProfile;
END_VAR
END_METHOD

METHOD PROF_GG_GERADE
VAR_INPUT
	PSCCHAR : POINTER TO L_MC2P_Characteristics;
	LRPOS : LREAL;
	PSCNORMSLAVE : POINTER TO L_MC2P_AxisProfile;
END_VAR
END_METHOD

METHOD PROF_GG_MODSIN
VAR_INPUT
	PSCCHAR : POINTER TO L_MC2P_Characteristics;
	LRPOS : LREAL;
	PSCNORMSLAVE : POINTER TO L_MC2P_AxisProfile;
END_VAR
END_METHOD

METHOD PROF_GG_POLY3
VAR_INPUT
	PSCCHAR : POINTER TO L_MC2P_Characteristics;
	LRPOS : LREAL;
	PSCNORMSLAVE : POINTER TO L_MC2P_AxisProfile;
END_VAR
END_METHOD

METHOD PROF_GR_POLY2
VAR_INPUT
	PSCCHAR : POINTER TO L_MC2P_Characteristics;
	LRPOS : LREAL;
	PSCNORMSLAVE : POINTER TO L_MC2P_AxisProfile;
END_VAR
END_METHOD

METHOD PROF_GU_HARMKOMB
VAR_INPUT
	PSCCHAR : POINTER TO L_MC2P_Characteristics;
	LRPOS : LREAL;
	PSCNORMSLAVE : POINTER TO L_MC2P_AxisProfile;
END_VAR
END_METHOD

METHOD PROF_RR_BESCHLTRAPEZ
VAR_INPUT
	PSCCHAR : POINTER TO L_MC2P_Characteristics;
	LRPOS : LREAL;
	PSCNORMSLAVE : POINTER TO L_MC2P_AxisProfile;
END_VAR
END_METHOD

METHOD PROF_RR_GENSIN
VAR_INPUT
	PSCCHAR : POINTER TO L_MC2P_Characteristics;
	LRPOS : LREAL;
	PSCNORMSLAVE : POINTER TO L_MC2P_AxisProfile;
END_VAR
END_METHOD

METHOD PROF_RR_MODBESCHLTRAPEZ
VAR_INPUT
	PSCCHAR : POINTER TO L_MC2P_Characteristics;
	LRPOS : LREAL;
	PSCNORMSLAVE : POINTER TO L_MC2P_AxisProfile;
END_VAR
END_METHOD

METHOD PROF_RR_QUADPARABEL
VAR_INPUT
	PSCCHAR : POINTER TO L_MC2P_Characteristics;
	LRPOS : LREAL;
	PSCNORMSLAVE : POINTER TO L_MC2P_AxisProfile;
END_VAR
END_METHOD

METHOD PROF_RR_SIN
VAR_INPUT
	PSCCHAR : POINTER TO L_MC2P_Characteristics;
	LRPOS : LREAL;
	PSCNORMSLAVE : POINTER TO L_MC2P_AxisProfile;
END_VAR
END_METHOD

METHOD PROF_RU_MODBESCHLTRAPEZ
VAR_INPUT
	PSCCHAR : POINTER TO L_MC2P_Characteristics;
	LRPOS : LREAL;
	PSCNORMSLAVE : POINTER TO L_MC2P_AxisProfile;
END_VAR
END_METHOD

METHOD PROF_UG_HARMKOMB
VAR_INPUT
	PSCCHAR : POINTER TO L_MC2P_Characteristics;
	LRPOS : LREAL;
	PSCNORMSLAVE : POINTER TO L_MC2P_AxisProfile;
END_VAR
END_METHOD

METHOD PROF_UR_MODBESCHLTRAPEZ
VAR_INPUT
	PSCCHAR : POINTER TO L_MC2P_Characteristics;
	LRPOS : LREAL;
	PSCNORMSLAVE : POINTER TO L_MC2P_AxisProfile;
END_VAR
END_METHOD

METHOD PROF_UU_SINGERKOMB
VAR_INPUT
	PSCCHAR : POINTER TO L_MC2P_Characteristics;
	LRPOS : LREAL;
	PSCNORMSLAVE : POINTER TO L_MC2P_AxisProfile;
END_VAR
END_METHOD

METHOD GETACCEQUIWITHA
END_METHOD

METHOD GETACCEQUIWITHOUTA
END_METHOD

METHOD GETACCNONEQUIWITHOUTA
END_METHOD

METHOD GETACCNONEQUIWITHA
END_METHOD

METHOD GETPOS
END_METHOD

METHOD GETVELEQUI
END_METHOD

METHOD GETVELNONEQUI
END_METHOD

(* ---- L_MC2P_CAMCREATOR.fb ---- *)
FUNCTION_BLOCK L_MC2P_CAMCREATOR
VAR_INPUT
	XENABLEINTERNALCAMTABLE : BOOL;
	XEXECUTE : BOOL;
	PCAMPOINTS : POINTER TO L_MC2P_CamDataXYVA;
	INUMOFPOINTS : INT;
	LRMASTERMAXVEL : LREAL;
	LRMASTERMAXACC : LREAL;
	LRMASTERSCALING : LREAL := 1;
	LRSLAVESCALING : LREAL := 1;
	SLAVE : AXIS_REF;
END_VAR
VAR_OUTPUT
	XINTERNALCAMTABLELACTIVE : BOOL;
	XERROR : BOOL;
	EERRORID : L_IE1P_Error;
	XBUSY : BOOL;
	XDONE : BOOL;
	CAMTABLEOUT : MC_CAM_REF;
	LRSLAVEMAXPOS : LREAL;
	LRSLAVEMINPOS : LREAL;
	LRSLAVEMAXVEL : LREAL;
	LRSLAVEMINVEL : LREAL;
	LRSLAVEMAXACC : LREAL;
	LRSLAVEMINACC : LREAL;
END_VAR
VAR
	EFMSTATE : L_MC2P_States := L_MC2P_States.INIT;
	SMC_CAMBOUNDS1 : L_MC2P_BoundsCam;
	CAMREF : L_MC2P_CamRefFromStruct;
	PCAMPOINTS_INT : POINTER TO L_MC2P_CamDataXYVA;
	INUMOFPOINTS_INT : INT;
	XINTERNALCONTROL : BOOL;
	XEXECUTE_OLD : BOOL;
	ASCCAMPOINTS : ARRAY [0..30] OF L_MC2P_CamDataXYVA;
	XINVALIDCAMTABLE : BOOL;
	XVISUACTIVE : BOOL := TRUE;
	DIFRAME : DINT;
	DIFRAME_OLD : DINT;
	ARVISPOINTLINES : ARRAY [1..10] OF L_MC2P_CamDataXYVA;
	IVISUTABLESETPOS : INT := 0;
	IVISUTABLESETPOS_OLD : INT := 0;
	IVISUTABLEMAXPOS : INT := 30;
	IVISSHOWLINESNO : INT;
	XVISPOINTMIN : BOOL;
	XVISPOINTMAX : BOOL;
	XVISUSETPOSUP : BOOL;
	XVISUSETPOSDOWN : BOOL;
	XVISUSETPOSUP_OLD : BOOL;
	XVISUSETPOSDOWN_OLD : BOOL;
	XSCROLBUTTENACTIVE : BOOL;
	TSETTIME : TIME := TIME#400ms;
	TON_SCROLBUTTEN : TON;
END_VAR
END_FUNCTION_BLOCK

METHOD CALL_CAMBOUNDS
END_METHOD

METHOD CALL_CAMREF
END_METHOD

METHOD CALL_CAMTABLEEQUIDISTANT
END_METHOD

METHOD CALL_CAMTABLENONEQUIDISTANT
END_METHOD

METHOD CALL_CAMTABLEPOLYNOMIAL
END_METHOD

METHOD CALL_ERRORHANDLER
END_METHOD

METHOD CALL_FBMETHODS
END_METHOD

METHOD CALL_INTERNALCTRL
END_METHOD

METHOD CALL_OUTPUT
END_METHOD

METHOD CALL_RESETCOMMANDS
END_METHOD

METHOD CALL_RESETOUTPUT
END_METHOD

METHOD CALL_STATEMACHINE
END_METHOD

METHOD CALL_VIS_TON_SCROLBUTTEN
END_METHOD

METHOD CALL_VISUTABCTRL
END_METHOD

METHOD CALL_VISUUPDATETAB
END_METHOD

METHOD DISABALE_VISU
END_METHOD

METHOD ENABLE_VISU
END_METHOD

METHOD CALL_S000_CYCLIC
END_METHOD

METHOD CALL_S001_INIT
END_METHOD

METHOD CALL_S002_READY
END_METHOD

(* ---- L_MC2P_CAMDATAOBJECT.fb ---- *)
FUNCTION_BLOCK L_MC2P_CAMDATAOBJECT
VAR_INPUT
	UCAMOBJECT : L_MC2P_XYVA;
	LRRESERVED : LREAL := 0;
END_VAR
VAR
	BASE : POINTER TO BYTE;
	DATATYPE : L_MC2P_MotionDataType;
	SIZE : UDINT;
	STARTADRESS : POINTER TO BYTE;
END_VAR
END_FUNCTION_BLOCK

(* ---- L_MC2P_CAMDATAPOINTXY.fb ---- *)
FUNCTION_BLOCK L_MC2P_CAMDATAPOINTXY
VAR_INPUT
	DWSTRUCTID : DWORD := L_MC2P_Constants.gC_dwCheckIDDataXY;
	LRX : LREAL;
	LRY : LREAL;
END_VAR
VAR
	BASE : POINTER TO BYTE;
	DATATYPE : L_MC2P_MotionDataType;
	SIZE : UDINT;
	STARTADRESS : POINTER TO BYTE;
END_VAR
END_FUNCTION_BLOCK

(* ---- L_MC2P_CAMDATAPOINTXYA.fb ---- *)
FUNCTION_BLOCK L_MC2P_CAMDATAPOINTXYA
VAR_INPUT
	DWSTRUCTID : DWORD := L_MC2P_Constants.gC_dwCheckIDDataXYA;
	LRX : LREAL;
	LRY : LREAL;
	LRYSS : LREAL;
END_VAR
VAR
	BASE : POINTER TO BYTE;
	DATATYPE : L_MC2P_MotionDataType;
	SIZE : UDINT;
	STARTADRESS : POINTER TO BYTE;
END_VAR
END_FUNCTION_BLOCK

(* ---- L_MC2P_CAMDATAPOINTY.fb ---- *)
FUNCTION_BLOCK L_MC2P_CAMDATAPOINTY
VAR_INPUT
	DWSTRUCTID : DWORD := L_MC2P_Constants.gC_dwCheckIDDataY;
	LRY : LREAL;
END_VAR
VAR
	BASE : POINTER TO BYTE;
	DATATYPE : L_MC2P_MotionDataType;
	SIZE : UDINT;
	STARTADRESS : POINTER TO BYTE;
END_VAR
END_FUNCTION_BLOCK

(* ---- L_MC2P_CAMDATAPOINTYA.fb ---- *)
FUNCTION_BLOCK L_MC2P_CAMDATAPOINTYA
VAR_INPUT
	DWSTRUCTID : DWORD := L_MC2P_Constants.gC_dwCheckIDDataYA;
	LRY : LREAL;
	LRYSS : LREAL;
END_VAR
VAR
	BASE : POINTER TO BYTE;
	DATATYPE : L_MC2P_MotionDataType;
	SIZE : UDINT;
	STARTADRESS : POINTER TO BYTE;
END_VAR
END_FUNCTION_BLOCK

(* ---- L_MC2P_CAMDATAXYVA.fb ---- *)
FUNCTION_BLOCK L_MC2P_CAMDATAXYVA
VAR_INPUT
	DWSTRUCTID : DWORD := L_MC2P_Constants.gC_dwCheckIDCond;
	ELAWOFMOTION : L_MC2P_LawOfMotion;
	LRX : LREAL;
	LRY : LREAL;
	LRYS : LREAL;
	LRYSS : LREAL;
	LRYSSS : LREAL;
	LRLAMBDA : LREAL := 0.5;
	LRPARAM1 : LREAL;
	LRPARAM2 : LREAL;
	LRPARAM3 : LREAL;
	LRPARAM4 : LREAL;
END_VAR
VAR
	BASE : POINTER TO BYTE;
	DATATYPE : L_MC2P_MotionDataType;
	SIZE : UDINT;
	STARTADRESS : POINTER TO BYTE;
END_VAR
END_FUNCTION_BLOCK

(* ---- L_MC2P_CAMEXTENDEDBASE.fb ---- *)
FUNCTION_BLOCK L_MC2P_CAMEXTENDEDBASE
VAR_INPUT
	MASTER : L_MC1P_IAXIS_REF_MASTERVALUES;
	XENABLE : BOOL;
	XSYNCCAM : BOOL;
	XSYNCOUTINSTANT : BOOL;
	XDIRECTCHANGE : BOOL;
	SCCAMTABLE : MC_CAM_REF;
	XPERIODIC : BOOL;
	LRCYCSETMASTERPOS : LREAL;
	LRCYCSETMASTERVEL : LREAL;
	LRCYCSETMASTERACC : LREAL;
	LRSETSLAVEPOS : LREAL;
	LRSETSLAVEVEL : LREAL;
	LRSETSLAVEACC : LREAL;
	ESYNCMODE : L_MC2P_ClutchMode;
	ESYNCDIRECTION : L_MC2P_ClutchDirection;
	LRMASTERSYNCINDIST : LREAL;
	LRMASTERSYNCINPOS : LREAL;
	LRMASTERSYNCOUTDIST : LREAL;
	LRSLAVESYNCOUTPOS : LREAL;
	LRLOADMASTERPOS_INT : LREAL;
	LRSYNCINTIME : LREAL;
	LRSYNCOUTTIME : LREAL;
	LRSYNCOUTINSTANTDEC : LREAL;
	LRSYNCCAMVEL : LREAL;
	LRSYNCCAMACC : LREAL;
	LRSYNCCAMDEC : LREAL;
	LRSYNCCAMJERK : LREAL;
END_VAR
VAR_OUTPUT
	XBUSY : BOOL;
	XERROR : BOOL;
	EERRORID : L_IE1P_Error;
	XCAMSYNCHRONISED : BOOL;
	XACCDECSYNC : BOOL;
	XENDOFPROFILE : BOOL;
	LRSETSLAVEPOSOUT : LREAL;
	LRSETSLAVEVELOUT : LREAL;
	LRSETSLAVEACCOUT : LREAL;
END_VAR
VAR_IN_OUT
	SLAVE : AXIS_REF;
END_VAR
VAR
	CLUTCHBASIC : L_MC2P_ClutchBasic;
	ESTATE : L_MC2P_States := L_MC2P_States.INIT;
	XSTATEENTRY : BOOL;
	XSMACTIVE : BOOL;
	XDONE : BOOL;
	XCONTINUOUSCAM_INT : BOOL;
	XNEWCAMTABLE : BOOL;
	XMASTEROUTOFSCALE : BOOL := FALSE;
	XINVALIDXVALUE : BOOL;
	XINVALIDSTARTENDVALUES : BOOL;
	XDIRECTCHANGE_INT : BOOL;
	SCCAMTABLE_INT : MC_Cam_REF;
	SCCAMINFO_INT : L_MC2P_CamInfo;
	XNOISEDETECTION_INT : BOOL := TRUE;
	LRTASKCYCLE_INT : LREAL;
	XPERIODIC_INT : BOOL;
	IENDOFPROFILECORECTION : INT;
	XNEXTAXISLIMIT : BOOL;
	LRCAMXSTART : LREAL;
	LRCAMXEND : LREAL;
	LRCAMXSTART_OLD : LREAL;
	LRCAMXEND_OLD : LREAL;
	LRCAMYSTART : LREAL;
	LRCAMYSTART_OLD : LREAL;
	LRCAMYEND : LREAL;
	LRCAMYEND_OLD : LREAL;
	ECAMPROFILER_CLUTCHMODE : L_MC2P_ClutchBasicMode;
	XSYNCOUTINSTANT_INT : BOOL;
	ESYNCDIRECTION_INT : L_MC2P_ClutchDirection;
	LRMASTERSYNCINDIST_INT : LREAL;
	LRMASTERSYNCINPOS_INT : LREAL;
	LRMASTERSYNCOUTDIST_INT : LREAL;
	LRSLAVESYNCOUTPOS_INT : LREAL;
	LRSYNCINTIME_INT : LREAL;
	LRSYNCOUTTIME_INT : LREAL;
	LRSYNCOUTINSTANTDEC_INT : LREAL;
	XSYNCCAM_OLD : BOOL;
	XENABLE_OLD : BOOL;
	XDIRECTCHANGE_OLD : BOOL;
	XSYNCOUTINSTANT_OLD : BOOL;
	LRCYCSETMASTERPOS_OLD : LREAL;
	LRSETXPOS_OLD : LREAL;
	XENDOFPROFILE_OLD : BOOL;
	XENDOFPROFPOSITIVE : BOOL;
	XENDOFPROFNEGATIVE : BOOL;
	LRENDOFPROFVARIANCE : LREAL := 1E-06;
	SCSETXPROFILE : L_MC2P_AxisProfile;
	SCSTARTYPROFILE : L_MC2P_AxisProfile;
	SCACTYPROFILE : L_MC2P_AxisProfile;
	SCACTYPROFILE_OLD : L_MC2P_AxisProfile;
	SCPROFGENXPROFILE : L_MC2P_AxisProfile;
	SCPROFGENYPROFILE : L_MC2P_AxisProfile;
	XCAMPROFILE_EXECUTE : BOOL;
	XCAMPROFILER_BUSY : BOOL;
	XCAMPROFILER_DONE : BOOL;
	XCAMPROFILER_INSYNC : BOOL;
	XCAMPROFILER_XACCDECSYNC : BOOL;
	XCAMPROFILER_XACCDECSYNC_OLD : BOOL;
	XCAMPROFILER_WARNINGCANTPREVENTREVERSE : BOOL;
	XCAMPROFILER_ERROR : BOOL;
	ECAMPROFILER_ERRORID : L_IE1P_Error;
	XCAMPROFILE_EXECUTE_OLD : BOOL;
	XFIRSTCYCLE : BOOL := TRUE;
	XEXTRAPOLATECAM : BOOL;
	XSTARTYPROFILECHECK : BOOL;
	LRSTARTYPROFILEMASTERDIST : LREAL;
	ALRMASTERPODDIFF : ARRAY [0..5] OF LREAL;
	FB_NOISEDETECTION : L_MC1P_NoiseDetection;
	FB_STACKVEL : L_MC1P_StackControlArray := STRUCT(iMaxLegth := 10);
	ALRVEL : ARRAY [1..10] OF LREAL;
	LRSUMVEL : LREAL;
	LRFILTMASTERVEL : LREAL;
	STARTINCURRENTPERIOD : BOOL;
	XNOISEDETECTION : BOOL;
END_VAR
END_FUNCTION_BLOCK

METHOD CALL_CAMPROFILER
END_METHOD

METHOD CALL_CHANGECAMTABLE_ENDOFPROFILE
END_METHOD

METHOD CALL_CHANGECAMTABLE_INSTANT
END_METHOD

METHOD CALL_CLUTCHCLOSEMODE
END_METHOD

METHOD CALL_CLUTCHOPENMODE
END_METHOD

METHOD CALL_CONVERTMASTERTOX
END_METHOD

METHOD CALL_CONVERTYTOSLAVE
END_METHOD

METHOD CALL_ERRORHANDLER
END_METHOD

METHOD CALL_FBMETHODS
END_METHOD

METHOD CALL_FB_NOISEDETECTION
END_METHOD

METHOD CALL_FIRSTCYCLE
END_METHOD

METHOD CALL_OUTPUT
END_METHOD

METHOD CALL_OUTPUT_ENDOFPROFILE
END_METHOD

METHOD CALL_RELEASECAM
VAR_INPUT
	SCOLDCAMTABLE : MC_Cam_REF;
END_VAR
END_METHOD

METHOD CALL_RESETCOMMANDS
END_METHOD

METHOD CALL_RESETOUTPUT
END_METHOD

METHOD CALL_STATEMASHINE
END_METHOD

METHOD CALL_STORECAMXYOLDVALUES
END_METHOD

METHOD SETPARCLUTCHCLOSE
END_METHOD

METHOD SETPARCLUTCHOPEN
END_METHOD

METHOD CALC_ENDOFPROFILEVALUES
END_METHOD

METHOD CALC_RESTARTSLAVEREL
END_METHOD

METHOD CALC_STARTYPROFILE
END_METHOD

METHOD CALC_XAXIS
END_METHOD

METHOD CALC_YAXIS
END_METHOD

METHOD CALL_RESETPROFGEN
END_METHOD

METHOD CAMTABLECHANGED : BOOL
VAR_INPUT
	SCCAMNEW : MC_Cam_REF;
	SCCAMOLD : MC_Cam_REF;
	SCCAMINFOOLD : L_MC2P_CamInfo;
END_VAR
END_METHOD

METHOD CAMTABLEVALID : BOOL
VAR_INPUT
	SCCAMTABLE : MC_Cam_REF;
END_VAR
END_METHOD

METHOD CHECK_XENDOFPERIOD : BOOL
VAR_OUTPUT
	XPOSITIVE : BOOL;
	XNEGATIVE : BOOL;
END_VAR
END_METHOD

METHOD COPYCAMTABLE
END_METHOD

METHOD FUN_AVERAGEMASTERVELFILTER : LREAL
VAR_INPUT
	XAVERAGEFILTER : BOOL;
	LRCYCMASTERVEL : LREAL;
END_VAR
END_METHOD

METHOD GET_INTERNCAMTABLE : MC_Cam_REF
END_METHOD

METHOD GET_ESTATE : L_MC2P_States
END_METHOD

METHOD GET_LRCAMPROFILERPOSOUT : LREAL
END_METHOD

METHOD GET_LRCAMXEND : LREAL
END_METHOD

METHOD GET_LRCAMXSTART : LREAL
END_METHOD

METHOD GET_LRCAMYEND : LREAL
END_METHOD

METHOD GET_LRCAMYSTART : LREAL
END_METHOD

METHOD GET_XCRITICALCYCLE : BOOL
END_METHOD

METHOD GET_XDONE : BOOL
END_METHOD

METHOD SET_ENDOFPROFVARIANCE
VAR_INPUT
	LRIN : LREAL;
END_VAR
END_METHOD

METHOD SET_INIT
END_METHOD

METHOD SET_INTERNCAMTABLE
VAR_INPUT
	CAMREF : MC_Cam_REF;
END_VAR
END_METHOD

METHOD CALL_S000_CYCLIC
END_METHOD

METHOD CALL_S001_INIT
END_METHOD

METHOD CALL_S002_CAM_DONE
END_METHOD

METHOD CALL_S010_01_READY_ENTRY_STATE
END_METHOD

METHOD CALL_S010_READY
END_METHOD

METHOD CALL_S100_CLUTCH_CLOSE
END_METHOD

METHOD CALL_S200_CAMMING
END_METHOD

METHOD CALL_S300_CLUTCH_OPEN
END_METHOD

METHOD CALL_S998_ERROR
END_METHOD

(* ---- L_MC2P_CAMEXTENDEDSTATE.fb ---- *)
FUNCTION_BLOCK L_MC2P_CAMEXTENDEDSTATE EXTENDS L_MC2P_CamExtendedBase
VAR_INPUT
	EOFFSETMODEMASTER : L_MC2P_OffsetMode;
	LRSETOFFSETMASTER : LREAL := 0.0;
	ESCALINGMODEMASTER : L_MC2P_ScalingMode;
	LRSETSCALINGMASTER : LREAL := 1.0;
	EOFFSETMODESLAVE : L_MC2P_OffsetMode;
	LRSETOFFSETSLAVE : LREAL := 0.0;
	ESCALINGMODESLAVE : L_MC2P_ScalingMode;
	LRSETSCALINGSLAVE : LREAL := 1.0;
	XMASTERABSOLUTE : BOOL;
	XSLAVEABSOLUTE : BOOL;
END_VAR
VAR_OUTPUT
	LRSETXPOSOUT : LREAL;
	LRSETXVELOUT : LREAL;
	LRSETXACCOUT : LREAL;
	LRSETYPOSOUT : LREAL;
	LRSETYVELOUT : LREAL;
	LRSETYACCOUT : LREAL;
END_VAR
VAR
	CAMAXISCONVERTER : L_MC2P_CamAxisConverter;
	EOFFSETMODEMASTER_INT : L_MC2P_OffsetMode;
	ESCALINGMODEMASTER_INT : L_MC2P_ScalingMode;
	XMASTERABSOLUTE_INT : BOOL;
	LRSETOFFSETMASTER_INT : LREAL;
	LRSETSCALINGMASTER_INT : LREAL;
	LRSETOFFSETMASTER_OLD : LREAL;
	LRSETOFFSETMASTER_2OLD : LREAL;
	LRSETOFFSETMASTER_3OLD : LREAL;
	XXAXISVALID : BOOL;
	ESCALINGMODESLAVE_INT : L_MC2P_ScalingMode;
	EOFFSETMODESLAVE_INT : L_MC2P_OffsetMode;
	LRSETOFFSETSLAVE_INT : LREAL;
	LRSETOFFSETSLAVE_OLD : LREAL;
	LRSETOFFSETSLAVE_2OLD : LREAL;
	LRSETSCALINGSLAVE_OLD : LREAL;
	LRSETSCALINGSLAVE_INT : LREAL;
	XLOADSLAVEPOSREL : BOOL;
	LRSETYPOSOUT_OLD : LREAL;
	LRTEMP : LREAL;
	SCACTYPROFILETEMP : L_MC2P_AxisProfile;
	SCPROFILETEMP : L_MC2P_AxisProfile;
	SCSETXPROFILETEMP : L_MC2P_AxisProfile;
	XMANIPULATEDXPOSFORENDOFPROFILE : BOOL;
	LRMASTERCYCLELENGTH : LREAL;
	LRMANIPULATEXPOSAFTERENDOFPROFILE : LREAL;
	XENDOFPROFPOSITIVE_INT : BOOL;
	XENDOFPROFNEGATIVE_INT : BOOL;
	XBLOCKCHECKENDOFPROFILE : BOOL;
	XOUTOFCAMPOSITIVE : BOOL;
	XOUTOFCAMNEGATIVE : BOOL;
	LRSETXPOSOUT_INT : LREAL;
	LRENDOFPROFILEWINDOW : LREAL;
	LRSETOFFSETVEL : LREAL;
	WSTARTYPROFILECHECKMODE : WORD := 0;
	WSTARTYPROFILECHECKMODE_RAMP_POS : WORD := 0;
	LWENDOFPROFILECHECKSUM : LWORD;
END_VAR
END_FUNCTION_BLOCK

METHOD CALL_CALCSLAVEAXISVALUES
END_METHOD

METHOD CALL_CALCXAXISVALUES
END_METHOD

METHOD CALL_CHANGECAMTABLE_ENDOFPROFILE
END_METHOD

METHOD CALL_CHANGECAMTABLE_INSTANT
END_METHOD

METHOD CALL_CONVERTMASTERTOX
END_METHOD

METHOD CALL_CONVERTYTOSLAVE
END_METHOD

METHOD CALL_ERRORHANDLER
END_METHOD

METHOD CALL_FBMETHODS
END_METHOD

METHOD CALL_OUTPUT
END_METHOD

METHOD CALL_PROFGENMASTER
END_METHOD

METHOD CALL_PROFGENSLAVE
END_METHOD

METHOD CALL_RESETAXISCONVERTER
END_METHOD

METHOD CALL_RESETCOMMANDS
END_METHOD

METHOD CALL_RESETOUTPUT
END_METHOD

METHOD CALL_SETMASTEROFFSET
END_METHOD

METHOD CALL_SETMASTERSCALING
END_METHOD

METHOD CALL_SETSLAVEOFFSET
END_METHOD

METHOD CALL_SETSLAVESCALING
END_METHOD

METHOD SETPARCLUTCHOPEN
END_METHOD

METHOD CALCCAMDATA : BOOL
END_METHOD

METHOD CALC_RESTARTSLAVEREL
END_METHOD

METHOD CALC_RESTARTXAXIS
END_METHOD

METHOD CALC_RESTARTYAXIS
END_METHOD

METHOD CALC_STARTYPROFILE
END_METHOD

METHOD CALC_XAXIS
END_METHOD

METHOD CALC_YAXIS
END_METHOD

METHOD CALC_LRSETOFFSETACCOUT : LREAL
VAR_IN_OUT
	LROFFSET : LREAL;
	LROFFSET_OLD : LREAL;
	LROFFSET_2OLD : LREAL;
	LRTASKCYCLE : LREAL;
END_VAR
END_METHOD

METHOD CALC_LRSETOFFSETVELOUT : LREAL
VAR_IN_OUT
	LROFFSET : LREAL;
	LROFFSET_OLD : LREAL;
	LRTASKCYCLE : LREAL;
END_VAR
END_METHOD

METHOD CALL_CORRECTIONMASTEROFFSETOLDVALUES
END_METHOD

METHOD CALL_MANIPULATEXPOSAFTERENDOFPROFILE : BOOL
END_METHOD

METHOD CALL_MANIPULATEYPOSAFTERENDOFPROFILE : BOOL
END_METHOD

METHOD CALL_RESETCAMBASIC
END_METHOD

METHOD CALL_RESETPROFGEN
END_METHOD

METHOD CHECK_XENDOFPERIOD : BOOL
VAR_OUTPUT
	XPOSITIVE : BOOL;
	XNEGATIVE : BOOL;
END_VAR
END_METHOD

METHOD CHECK_XENDOFPERIODBEFORCAMPROFILER : BOOL
END_METHOD

METHOD GET_LRACTIVESCALINGMASTER : LREAL
END_METHOD

METHOD GET_LRACTIVESCALINGSLAVE : LREAL
END_METHOD

METHOD GET_LRCONVERTMASTERTOXPOS : LREAL
END_METHOD

METHOD GET_LRCONVERTYTOSLAVEPOS : LREAL
END_METHOD

METHOD GET_LRSETY : LREAL
END_METHOD

METHOD GET_LRSLAVEOFFSETREL : LREAL
END_METHOD

METHOD GET_LRXOFFSETREL : LREAL
END_METHOD

METHOD GET_XENDOFPROFNEGATIVE : BOOL
END_METHOD

METHOD GET_XENDOFPROFPOSITIVE : BOOL
END_METHOD

METHOD SET_LRENDOFPROFILEFACTOR : BOOL
VAR_INPUT
	LRIN : LREAL := 1;
END_VAR
END_METHOD

METHOD SET_LRENDOFPROFILEWINDOW : BOOL
VAR_INPUT
	LRIN : LREAL := 1;
END_VAR
END_METHOD

METHOD CALL_S000_CYCLIC
END_METHOD

METHOD CALL_S001_INIT
END_METHOD

METHOD CALL_S002_CAM_DONE
END_METHOD

METHOD CALL_S010_01_READY_ENTRY_STATE
END_METHOD

METHOD CALL_S998_ERROR
END_METHOD

(* ---- L_MC2P_CAMGETSLAVEPOSITION.fb ---- *)
FUNCTION_BLOCK L_MC2P_CAMGETSLAVEPOSITION EXTENDS L_MC2P_CamBasic
VAR_INPUT
	XEXECUTE : BOOL;
	LRMASTERPOSITION : LREAL;
	ITFCAMTABLE : MC_CAM_REF;
END_VAR
VAR_OUTPUT
	XDONE : BOOL;
	XBUSY : BOOL;
	XERROR : BOOL;
	EERRORID : L_IE1P_Error;
	LRSLAVEPOSITION : LREAL;
END_VAR
VAR
	SCINPUTMASTER_INT : L_MC2P_AxisProfile;
	SCOUTPUTSLAVE_INT : L_MC2P_AxisProfile;
	XEXECUTEOLD : BOOL;
END_VAR
END_FUNCTION_BLOCK

(* ---- L_MC2P_CAMREFFROMFILE.fb ---- *)
FUNCTION_BLOCK L_MC2P_CAMREFFROMFILE EXTENDS L_MC2P_ReadLMDFile
VAR_INPUT
	XEXECUTE : BOOL;
	SFILENAME : STRING := '';
	ITFCAMDATA : L_MC2P_IMotionData;
	UDICAMDATACOUNT : UDINT;
	XRELOADABLE : BOOL;
END_VAR
VAR_OUTPUT
	XDONE : BOOL;
	XBUSY : BOOL;
	XERROR : BOOL;
	EERRORID : L_IE1P_Error;
END_VAR
VAR
	MOTIONDATA_INT : L_MC2P_IMotionData;
	SCCAMDATA : L_MC2P_CamData;
	XRELOADOLD : BOOL;
	STEMPFILE : STRING;
	RELOAD : BOOL;
END_VAR
END_FUNCTION_BLOCK

METHOD CHECKFILENAME : BOOL
VAR_IN_OUT
	SFILE : STRING;
END_VAR
END_METHOD

METHOD CHECKINPUTS : BOOL
END_METHOD

METHOD LOADDATA
END_METHOD

METHOD MAIN
END_METHOD

METHOD GETCAMDATA : POINTER TO L_MC2P_CamData
END_METHOD

METHOD GETID : DWORD
END_METHOD

METHOD SETCAMDATAACTIVE
VAR_INPUT
	XCAMACITVE : BOOL;
END_VAR
END_METHOD

METHOD SETMASTERVALUES
VAR_INPUT
	LRMASTERPOS : LREAL;
END_VAR
END_METHOD

METHOD GETCOND
VAR_INPUT
	HFILE : SYSFILE.RTS_IEC_HANDLE;
	ITFCAMDATA : L_MC2P_IMotionData;
	WDATAELEMENTS : WORD;
	DWCOUNT : DWORD;
END_VAR
END_METHOD

METHOD GETDATAPOINTS
VAR_INPUT
	HFILE : SYSFILE.RTS_IEC_HANDLE;
	ITFCAMDATA : L_MC2P_IMotionData;
	WDATAELEMENTS : WORD;
	DWCOUNT : DWORD;
	XWITHPRECONTROL : BOOL;
END_VAR
END_METHOD

METHOD READCAMDATA
VAR_INPUT
	HFILE : SYSFILE.RTS_IEC_HANDLE;
END_VAR
END_METHOD

METHOD READSPECIFICDATA
VAR_INPUT
	HFILE : SYSFILE.RTS_IEC_HANDLE;
END_VAR
END_METHOD

(* ---- L_MC2P_CAMREFFROMSTRUCT.fb ---- *)
FUNCTION_BLOCK L_MC2P_CAMREFFROMSTRUCT EXTENDS L_MC2P_TemplateNoAxis
VAR_INPUT
	XEXECUTE : BOOL;
	SNAME : STRING(50);
	UDICAMDATACOUNT : UDINT;
	ITFCAMDATA : L_MC2P_IMotionData;
	ECAMTYPE : L_MC2P_CamType;
	EINTERPOLATIONQUALITY : L_MC2P_InterpolationQuality;
	LRXSTARTPOS : LREAL;
	LRXENDPOS : LREAL;
END_VAR
VAR_OUTPUT
	XDONE : BOOL;
	XBUSY : BOOL;
	XERROR : BOOL;
	EERRORID : L_IE1P_Error;
END_VAR
VAR
	I : UDINT;
	SCCAMDATA : L_MC2P_CamData;
	PCAMDATAXYVA : POINTER TO L_MC2P_CamDataXYVA;
	PCAMDATAPOINTXYA : POINTER TO L_MC2P_CamDataPointXYA;
	PCAMDATAPOINTXY : POINTER TO L_MC2P_CamDataPointXY;
	PCAMDATAPOINTY : POINTER TO L_MC2P_CamDataPointY;
	PCAMDATAPOINTYA : POINTER TO L_MC2P_CamDataPointYA;
	XEXECUTEOLD : BOOL;
	XRESETOUTPUT : BOOL;
	XDATAVALID : BOOL;
	XDATAACTIVE : BOOL;
	DWDATACRC : DWORD;
	LRACTXPOS : LREAL;
END_VAR
END_FUNCTION_BLOCK

METHOD GETCAMDATA : POINTER TO L_MC2P_CamData
END_METHOD

METHOD GETID : DWORD
END_METHOD

METHOD SETCAMDATAACTIVE
VAR_INPUT
	XCAMACITVE : BOOL;
END_VAR
END_METHOD

METHOD SETMASTERVALUES
VAR_INPUT
	LRMASTERPOS : LREAL;
END_VAR
END_METHOD

(* ---- L_MC2P_CAMREFTOFILE.fb ---- *)
FUNCTION_BLOCK L_MC2P_CAMREFTOFILE EXTENDS L_MC2P_WriteLMDFile
VAR_INPUT
	XEXECUTE : BOOL;
	SFILENAME : STRING := '';
	ITFCAMTABLE : MC_CAM_REF;
END_VAR
VAR_OUTPUT
	XDONE : BOOL;
	XBUSY : BOOL;
	XERROR : BOOL;
	EERRORID : L_IE1P_Error;
END_VAR
VAR
	XRELOADOLD : BOOL;
	RELOAD : BOOL;
END_VAR
END_FUNCTION_BLOCK

METHOD MAIN
END_METHOD

METHOD WRITECAMDATA
VAR_INPUT
	HFILE : SYSFILE.RTS_IEC_HANDLE;
END_VAR
END_METHOD

METHOD WRITECOND
VAR_INPUT
	HFILE : SYSFILE.RTS_IEC_HANDLE;
	ITFCAMDATA : L_MC2P_IMotionData;
	DWCOUNT : DWORD;
END_VAR
END_METHOD

METHOD WRITEDATAPOINTS
VAR_INPUT
	HFILE : SYSFILE.RTS_IEC_HANDLE;
	ITFCAMDATA : L_MC2P_IMotionData;
	DWCOUNT : DWORD;
	XWITHPRECONTROL : BOOL;
END_VAR
END_METHOD

METHOD WRITESPECIFICDATA
VAR_INPUT
	HFILE : SYSFILE.RTS_IEC_HANDLE;
END_VAR
END_METHOD

(* ---- L_MC2P_CAMTABLEINFO.fb ---- *)
FUNCTION_BLOCK L_MC2P_CAMTABLEINFO
VAR_INPUT
	XENABLE : BOOL;
	CAMTABLE : MC_CAM_REF;
	LRMASTERMAXVEL : LREAL := 100;
	LRMASTERMAXACC : LREAL := 1000;
	LRMASTERSCALING : LREAL := 1;
	LRSLAVESCALING : LREAL := 1;
END_VAR
VAR_OUTPUT
	XBUSY : BOOL;
	XDONE : BOOL;
	XCAMTABLEVALID : BOOL;
	LRMASTERSTARTPOS : LREAL;
	LRMASTERENDPOS : LREAL;
	LRSLAVESTARTPOS : LREAL;
	LRSLAVEENDPOS : LREAL;
	LRSLAVEMAXPOS : LREAL;
	LRSLAVEMINPOS : LREAL;
	LRSLAVEMAXVEL : LREAL;
	LRSLAVEMINVEL : LREAL;
	LRSLAVEMAXACC : LREAL;
	LRSLAVEMINACC : LREAL;
END_VAR
VAR
	EFMSTATE : L_MC2P_States := L_MC2P_States.INIT;
	CAMTABLE_INT : MC_CAM_REF;
	XENABLE_OLD : BOOL;
	SMC_CAMBOUNDS1 : L_MC2P_BoundsCam;
	XCALCNEWVALUES : BOOL;
END_VAR
END_FUNCTION_BLOCK

METHOD CALC_STARTENDVALUES
END_METHOD

METHOD CALL_CAMBOUNDS
END_METHOD

METHOD CALL_FBMETHODS
END_METHOD

METHOD CALL_OUTPUT
END_METHOD

METHOD CALL_RESETCOMMANDS
END_METHOD

METHOD CALL_RESETOUTPUT
END_METHOD

METHOD CALL_STATEMACHINE
END_METHOD

METHOD GET_XCALCNEWVALUES : BOOL
END_METHOD

METHOD GET_XCRITICALCYCLE : BOOL
END_METHOD

METHOD CALL_S000_CYCLIC
END_METHOD

(* ---- L_MC2P_CLUTCHBASIC.fb ---- *)
FUNCTION_BLOCK L_MC2P_CLUTCHBASIC
VAR
	L_MC2P_CAMBASIC1 : L_MC2P_CamBasic;
	XBUSYMAIN : BOOL;
	XDONEMAIN : BOOL;
	XERRORMAIN : BOOL;
	EERRORIDMAIN : L_IE1P_Error;
	ECLUTCHMODEMAIN : WORD;
	XRESETOUTPUTMAIN : BOOL;
	XBUSYINT : BOOL;
	XBUSYINT2 : BOOL;
	XDONEINT : BOOL;
	XDONEINT2 : BOOL;
	XWARNINGCANTPREVENTREVERSEINT : BOOL;
	XERRORINT : BOOL;
	EERRORIDINT : L_IE1P_Error;
	XEXECUTEOLD : BOOL;
	XCLUTCHOLD : BOOL;
	XRESET : BOOL;
	XRESETOUTPUT : BOOL;
	XCLUTCHACC : BOOL;
	LRENDTIME : LREAL;
	SCSLAVEEND : L_MC2P_AxisProfile;
	SCSLAVESTART : L_MC2P_AxisProfile;
	SCMASTEREND : L_MC2P_AxisProfile;
	SCMASTERSTART : L_MC2P_AxisProfile;
	UDICOUNTER : UDINT;
	LRPOSOLD : LREAL;
	LRVELOLD : LREAL;
	XFLAGCLUTCH : BOOL;
	LRMASTERSTART_INT : LREAL;
	LRMASTEREND_INT : LREAL;
	LRSLAVESTART_INT : LREAL;
	LRSLAVEEND_INT : LREAL;
	XREVERSEALLOWED : BOOL;
	XREDUCEACC : BOOL;
	XCHECKREVERSEBEFORECLUTCH : BOOL;
	LROLDMAPOS : LREAL;
	LRMASTERSTARTPOSITION : LREAL;
	LRMASTERENDPOSITION : LREAL;
	LRMASTERCLUTCHPOSITION_INT : LREAL;
	LRMASTERCLUTCHDISTANCE_INT : LREAL;
	LRMASTEROPENPOS : LREAL;
	SCCHARCLUTCH : ARRAY [0..1] OF L_MC2P_Characteristics;
	ICORRECT : INT;
	ICLUTCHSTARTCOUNTER : INT;
	XCLUTCHSTARTFORWARD : BOOL;
	XCLUTCHSTARTBACKWARD : BOOL;
	XCLUTCHSTARTFORWARDSET : BOOL;
	XCLUTCHSTARTBACKWARDSET : BOOL;
	XCLUTCHREADYFORWARD : BOOL;
	XCLUTCHREADYBACKWARD : BOOL;
	XCLUTCHREADY : BOOL;
	XSETSTARTPOS : BOOL;
	XDIRECTIONSTARTPOS : BOOL;
	PG : L_MC1P_PosProfiler;
	SCPARAM : L_MC1P_ProfileParameter;
	XPOSMODE : BOOL;
	RG : L_MC1P_RampGeneratorIntern;
	LRMAPOSOLDMAIN : LREAL;
	XCORRECTCLUTCHOFFSETNEXTCYCLE : BOOL;
	XCORRECTCLUTCHOFFSETACTCYCLE : BOOL;
	LRCLUTCHOFFSET : LREAL;
	LRJERKSET : LREAL;
	LRSAVEPOS : LREAL;
	LRSAVEVEL : LREAL;
	XSYNCINOUTOLD : BOOL;
	XWAITSTART : BOOL;
	XSTARTINCURRENTPERIOD : BOOL := FALSE;
	EACTMASTERDIRECTION : L_MC2P_Direction;
	EACTMASTERDIRECTIONOLD : L_MC2P_Direction;
	LRMAXNOISE : LREAL;
	LRMINNOISE : LREAL;
	XUPDATESETVALUEFIRSTCLUTCHCYCLE : BOOL;
	CHARCLUTCH : ARRAY [0..1] OF L_MC2P_Characteristics;
	CLUTCHOFFSET : LREAL;
	CORRECTCLUTCHOFFSETACTCYCLE : BOOL;
	CORRECTCLUTCHOFFSETNEXTCYCLE : BOOL;
	MASTERDIRECTION : L_MC2P_Direction;
	STARTINCURRENTPERIOD : BOOL;
	UPDATESETVALUEFIRSTCLUTCHCYCLE : BOOL;
END_VAR
END_FUNCTION_BLOCK

METHOD CALCULATECOMPLETECAMPROFILE
VAR_INPUT
	XEXECUTE : BOOL;
	PCAMDATA : POINTER TO L_MC2P_CamData;
	SCINPUTMASTER : L_MC2P_AxisProfile;
	SCACTSLAVE : L_MC2P_AxisProfile;
	ECLUTCHMODE : L_MC2P_ClutchBasicMode := 0;
	LRMASTERCLOSEDIST : LREAL;
	LRMASTERCLOSEPOS : LREAL;
	LRMASTEROPENDIST : LREAL;
	LRSLAVEOPENPOS : LREAL;
	LRLOADMASTERPOS : LREAL;
	EMASTERDIRECTION : L_MC2P_ClutchDirection := L_MC2P_ClutchDirection.mcCurrentDirection;
	LROPENTIME : LREAL;
	LRCLOSETIME : LREAL;
	LRCLOSEONTIMEOFFSET : LREAL;
	LRDECOPENINSTANT : LREAL;
	LRMAXVELDIFF : LREAL;
	LRMAXACC : LREAL;
	LRMAXDEC : LREAL;
	LRJERK : LREAL;
	LRCYCLETIME : LREAL;
	LRJERKDEFAULT : LREAL;
	EMASTERAXISTYPE : L_MC1P_TraversingRange;
	XPERIODIC : BOOL;
	PSCOUTPUTSLAVE : POINTER TO L_MC2P_AxisProfile;
	XEXTRAPOLATECAM : BOOL;
END_VAR
VAR_OUTPUT
	XBUSY : BOOL;
	XDONE : BOOL;
	XINSYNC : BOOL;
	XCLUTCHACTIVE : BOOL;
	XWARNINGCANTPREVENTREVERSE : BOOL;
	XERROR : BOOL;
	EERRORID : L_IE1P_Error;
END_VAR
END_METHOD

METHOD CHECKPOSNOISE
VAR_IN_OUT
	LRCYCPOS : LREAL;
	LRCYCLELENGTH : LREAL;
END_VAR
END_METHOD

METHOD CLOSEONLIMITED
VAR_INPUT
	XCLUTCH : BOOL;
	SCINPUTSLAVE : L_MC2P_AxisProfile;
	SCACTSLAVE : L_MC2P_AxisProfile;
	XPOSMODE : BOOL;
	LRMAXVELDIFF : LREAL;
	LRMAXACC : LREAL;
	LRMAXDEC : LREAL;
	LRJERK : LREAL;
	LRCYCLETIME : LREAL;
END_VAR
VAR_OUTPUT
	SCOUTPUTSLAVE : L_MC2P_AxisProfile;
	XBUSY : BOOL;
	XDONE : BOOL;
	XERROR : BOOL;
	EERRORID : L_IE1P_Error;
END_VAR
END_METHOD

METHOD CLOSEONSPEED
VAR_INPUT
	XCLUTCH : BOOL;
	SCINPUTSLAVE : L_MC2P_AxisProfile;
	SCACTSLAVE : L_MC2P_AxisProfile;
	LRMAXACC : LREAL;
	LRMAXDEC : LREAL;
	LRJERK : LREAL;
	LRCYCLETIME : LREAL;
END_VAR
VAR_OUTPUT
	SCOUTPUTSLAVE : L_MC2P_AxisProfile;
	XBUSY : BOOL;
	XDONE : BOOL;
	XERROR : BOOL;
	EERRORID : L_IE1P_Error;
END_VAR
END_METHOD

METHOD CLOSEONTIME
VAR_INPUT
	XCLUTCH : BOOL;
	SCINPUTSLAVE : L_MC2P_AxisProfile;
	SCACTSLAVE : L_MC2P_AxisProfile;
	LRCLOSETIME : LREAL := 0.001;
	LRCYCLETIME : LREAL := 0.001;
END_VAR
VAR_OUTPUT
	SCOUTPUTSLAVE : L_MC2P_AxisProfile;
	XBUSY : BOOL;
	XDONE : BOOL;
	XERROR : BOOL;
	EERRORID : L_IE1P_Error;
END_VAR
END_METHOD

METHOD CLUTCHONPOSITION
VAR_INPUT
	XCLUTCH : BOOL;
	SCINPUTMASTER : L_MC2P_AxisProfile;
	SCSLAVEACT : L_MC2P_AxisProfile;
	SCSLAVEEND : L_MC2P_AxisProfile;
	LRMASTERCLUTCHPOSITION : LREAL;
	LRMASTERCLUTCHDISTANCE : LREAL;
	EMASTERDIRECTION : L_MC2P_ClutchDirection;
	LRMASTERSTARTPOS : LREAL;
	LRMASTERENDPOS : LREAL;
	LRSLAVESTARTPOS : LREAL;
	LRSLAVEENDPOS : LREAL;
	LRCYCLETIME : LREAL;
	EMASTERAXISTYPE : L_MC1P_TraversingRange;
	XREVERSEALLOWED : BOOL;
	XCLUTCHSLAVE : BOOL;
	XPERIODIC : BOOL;
	LRJERK : LREAL;
END_VAR
VAR_OUTPUT
	SCOUTPUTSLAVE : L_MC2P_AxisProfile;
	XBUSY : BOOL;
	XCLUTCHACTIVE : BOOL;
	XDONE : BOOL;
	XERROR : BOOL;
	EERRORID : L_IE1P_Error;
END_VAR
END_METHOD

METHOD CLUTCHONPOSITION_2
VAR_INPUT
	XCLUTCH : BOOL;
	SCINPUTMASTER : L_MC2P_AxisProfile;
	SCSLAVEACT : L_MC2P_AxisProfile;
	SCSLAVEEND : L_MC2P_AxisProfile;
	LRMASTERCLUTCHPOSITION : LREAL;
	LRMASTERCLUTCHDISTANCE : LREAL;
	EMASTERDIRECTION : L_MC2P_ClutchDirection;
	LRMASTERSTARTPOS : LREAL;
	LRMASTERENDPOS : LREAL;
	LRSLAVESTARTPOS : LREAL;
	LRSLAVEENDPOS : LREAL;
	LRCYCLETIME : LREAL;
	EMASTERAXISTYPE : L_MC1P_TraversingRange;
	XREVERSEALLOWED : BOOL;
	XCLUTCHSLAVE : BOOL;
	XPERIODIC : BOOL;
	LRJERK : LREAL;
END_VAR
VAR_OUTPUT
	SCOUTPUTSLAVE : L_MC2P_AxisProfile;
	XBUSY : BOOL;
	XCLUTCHACTIVE : BOOL;
	XDONE : BOOL;
	XERROR : BOOL;
	EERRORID : L_IE1P_Error;
END_VAR
END_METHOD

METHOD GENERATECLUTCHONPOSITIONMASTER
VAR_INPUT
	SCACTMASTER : L_MC2P_AxisProfile;
	SCSTARTMASTER : L_MC2P_AxisProfile;
	SCENDMASTER : L_MC2P_AxisProfile;
	LRMASTERSTARTPOSITION : LREAL;
	LRMASTERCLUTCHPOSITION : LREAL;
	LRMASTERCLUTCHDISTANCE : LREAL;
	LRMASTERSTART : LREAL;
	PSCCHARCLUTCH : POINTER TO L_MC2P_Characteristics;
	XMASTERPOSITIVEDIRECTION : BOOL;
END_VAR
END_METHOD

METHOD GENERATECLUTCHONPOSITIONSLAVE
VAR_INPUT
	SCACTMASTER : L_MC2P_AxisProfile;
	SCSTARTSLAVE : L_MC2P_AxisProfile;
	SCENDSLAVE : L_MC2P_AxisProfile;
	LRMASTERSTARTPOSITION : LREAL;
	LRMASTERCLUTCHPOSITION : LREAL;
	LRMASTERCLUTCHDISTANCE : LREAL;
	LRMASTERSTART : LREAL;
	LRMASTEREND : LREAL;
	LRSLAVEPOSDIFF : LREAL;
	UINUMOFCYCLESMASTER : UINT;
	UINUMOFCYCLESSLAVE : UINT;
	PSCCHARCLUTCH : POINTER TO L_MC2P_Characteristics;
	EMASTERAXISTYPE : L_MC1P_TraversingRange;
	XMASTERPOSITIVEDIRECTION : BOOL;
END_VAR
END_METHOD

METHOD GENERATESYNCONPOSITION
VAR_INPUT
	XDIRECTIONPOSITIVE : BOOL;
	LRMASTERSTARTPOSITION : LREAL;
	LRMASTERENDPOSITION : LREAL;
	LRSLAVESTARTPOSITION : LREAL;
	LRSLAVEENDPOSITION : LREAL;
	XSYNCONSTART : BOOL;
	PSCCHARCLUTCH : POINTER TO L_MC2P_Characteristics;
END_VAR
END_METHOD

METHOD OPENINSTANT
VAR_INPUT
	XCLUTCH : BOOL;
	SCINPUTSLAVE : L_MC2P_AxisProfile;
	LRDECOPENINSTANT : LREAL;
	LRCYCLETIME : LREAL;
END_VAR
VAR_OUTPUT
	SCOUTPUTSLAVE : L_MC2P_AxisProfile;
	XBUSY : BOOL;
	XDONE : BOOL;
	XERROR : BOOL;
	EERRORID : L_IE1P_Error;
END_VAR
END_METHOD

METHOD OPENONCONSTVELOCITY
VAR_INPUT
	XCLUTCH : BOOL;
	SCINPUTSLAVE : L_MC2P_AxisProfile;
	LRMAXDEC : LREAL;
	LRJERK : LREAL;
	LRCYCLETIME : LREAL;
END_VAR
VAR_OUTPUT
	SCOUTPUTSLAVE : L_MC2P_AxisProfile;
	XBUSY : BOOL;
	XDONE : BOOL;
	XERROR : BOOL;
	EERRORID : L_IE1P_Error;
END_VAR
END_METHOD

METHOD OPENONLIMITED
VAR_INPUT
	XCLUTCH : BOOL;
	SCINPUTSLAVE : L_MC2P_AxisProfile;
	XPOSMODE : BOOL;
	LRSLAVEOPENPOS : LREAL;
	LRMAXVELDIFF : LREAL;
	LRMAXACC : LREAL;
	LRMAXDEC : LREAL;
	LRJERK : LREAL;
	LRCYCLETIME : LREAL;
END_VAR
VAR_OUTPUT
	SCOUTPUTSLAVE : L_MC2P_AxisProfile;
	XBUSY : BOOL;
	XDONE : BOOL;
	XERROR : BOOL;
	EERRORID : L_IE1P_Error;
END_VAR
END_METHOD

METHOD OPENONREDUCEACC
VAR_INPUT
	XCLUTCH : BOOL;
	SCACTSLAVE : L_MC2P_AxisProfile;
	XREVERSEALLOWED : BOOL;
	LRJERK : LREAL;
	LRCYCLETIME : LREAL;
END_VAR
VAR_OUTPUT
	SCOUTPUTSLAVE : L_MC2P_AxisProfile;
	XBUSY : BOOL;
	XDONE : BOOL;
	XWARNINGCANTPREVENTREVERSE : BOOL;
	XERROR : BOOL;
	EERRORID : L_IE1P_Error;
END_VAR
END_METHOD

METHOD OPENONTIME
VAR_INPUT
	XCLUTCH : BOOL;
	SCINPUTSLAVE : L_MC2P_AxisProfile;
	SCACTSLAVE : L_MC2P_AxisProfile;
	LRSLAVEOPENPOS : LREAL := 0;
	LROPENTIME : LREAL := 0.001;
	LRCYCLETIME : LREAL := 0.001;
END_VAR
VAR_OUTPUT
	SCOUTPUTSLAVE : L_MC2P_AxisProfile;
	XBUSY : BOOL;
	XDONE : BOOL;
	XERROR : BOOL;
	EERRORID : L_IE1P_Error;
END_VAR
END_METHOD

METHOD PROFILECLUTCHONPOSITION
VAR_INPUT
	SCACTMASTER : L_MC2P_AxisProfile;
	SCCHARCLUTCH : ARRAY [0..1] OF L_MC2P_Characteristics;
	LRMASTERSTART : LREAL;
	LRMASTEREND : LREAL;
	XSTARTCLUTCH : BOOL;
	EMASTERAXISTYPE : L_MC1P_TraversingRange;
	XMASTERPOSITIVEDIRECTION : BOOL;
END_VAR
VAR_OUTPUT
	SCACTSLAVE : L_MC2P_AxisProfile;
END_VAR
END_METHOD

METHOD PROFILESYNCONPOSITION : INT
VAR_INPUT
	SCACTMASTER : L_MC2P_AxisProfile;
	SCCHARCLUTCH : ARRAY [0..1] OF L_MC2P_Characteristics;
	LRMASTERSTARTPOSITION : LREAL;
	LRMASTERSTART : LREAL;
	LRMASTEREND : LREAL;
	XSTARTCLUTCH : BOOL;
	PSCACTSLAVE : POINTER TO L_MC2P_AxisProfile;
END_VAR
END_METHOD

METHOD RESETCLUTCH
END_METHOD

METHOD RESETSTARTFLAG
END_METHOD

METHOD SYNCONPOSITION
VAR_INPUT
	XSYNCINOUT : BOOL;
	XSYNCMODEIN : BOOL;
	SCINPUTMASTER : L_MC2P_AxisProfile;
	SCINPUTSLAVE : L_MC2P_AxisProfile;
	LRSYNCPOSITION : LREAL;
	LRSYNCDISTANCE : LREAL;
	LRMASTERSTARTPOS : LREAL;
	LRMASTERENDPOS : LREAL;
	LRSLAVESTARTPOS : LREAL;
	LRSLAVEENDPOS : LREAL;
	IMASTERMOVEMENTTYPE : INT;
	XPERIODIC : BOOL;
	PSCOUTPUTSLAVE : POINTER TO L_MC2P_AxisProfile;
END_VAR
VAR_OUTPUT
	XBUSY : BOOL;
	XCLUTCHACTIVE : BOOL;
	XDONE : BOOL;
	XWARNINGCANTPREVENTREVERSE : BOOL;
	XERROR : BOOL;
	EERRORID : L_IE1P_Error;
END_VAR
END_METHOD

(* ---- L_MC2P_CLUTCHPOS.fb ---- *)
FUNCTION_BLOCK L_MC2P_CLUTCHPOS
VAR_INPUT
	LRSETCYCPOS : LREAL;
	XOPEN : BOOL;
	LROPENPOSITION : LREAL;
	XOPENINSTANT : BOOL;
	XRESET : BOOL;
	LRDISTENGAGE : LREAL := 90;
	LRDISTDISENGAGE : LREAL := 90;
	LRDEC : LREAL;
	LRJERK : LREAL;
	ETRAVERSINGRANGE : L_MC1P_TraversingRange;
	LRCYCLELENGTH : LREAL;
END_VAR
VAR_OUTPUT
	LRSETPOSOUT : LREAL;
	LRSETVELOUT : LREAL;
	XCLOSED : BOOL;
	XOPENDONE : BOOL;
	XINTARGET : BOOL;
	XERROR : BOOL;
	EERRORID : L_IE1P_Error;
END_VAR
VAR
	LRTASKCYCLE : LREAL;
	NSTEPCOUNTER : INT;
	NACTION : INT;
	LRSAVEPOSIN : LREAL;
	LRDIFFIN : LREAL;
	LRVELRAMP : LREAL;
	LRINTEGRATOR : LREAL;
	LRSETPOS : LREAL;
	LRSTARTPOSITION : LREAL;
	LRENDPOSITION : LREAL;
	LRACTPOS : LREAL;
	LRSAVEPOSOUT : LREAL;
	LRDIFF : LREAL;
	LROPENPOS : LREAL;
	LRDIFFOPENINS : LREAL;
	NINDICATOR : INT;
	LRPOSINT : LREAL;
	RAMPGEN : L_MC1P_RampGeneratorIntern;
	LRCYCLELENINT : LREAL;
	INDICATOR_CW : INT := 20;
	INDICATOR_CCW : INT := -20;
	NOACTION : INT := 0;
	ENGAGE : INT := 1;
	DISENGAGE : INT := 2;
	CLUTCHP_CLOSE : INT := 0;
	CLUTCHP_OPEN_START_CW : INT := 2;
	CLUTCHP_OPEN_START_CCW : INT := 3;
	CLUTCHP_OPEN_DONE : INT := 5;
	CLUTCHP_CLOSE_START_CW : INT := 7;
	CLUTCHP_CLOSE_START_CCW : INT := 8;
	CLUTCHP_CLOSE_DONE : INT := 11;
	CLUTCHP_OPEN_WARNING : INT := 15;
	CLUTCHP_OPENINSTANT_START : INT := 16;
	CLUTCHP_OPENINSTANT_DONE : INT := 17;
	CLUTCHP_OPENINSTANT_QUIT : INT := 18;
END_VAR
END_FUNCTION_BLOCK

METHOD GETENDPOS : LREAL
VAR_INPUT
	LRSETVELOCITY : LREAL;
	LRSTARTPOSITION : LREAL;
	LRCLOSEDISTANCE : LREAL;
END_VAR
END_METHOD

METHOD GETENDPOSOPEN : LREAL
VAR_INPUT
	LRSETVELOCITY : LREAL;
	LRSTARTPOSITION : LREAL;
	LROPENPOSITION : LREAL;
	LROPENDISTANCE : LREAL;
	LRCYCLELENGTH : LREAL;
END_VAR
END_METHOD

METHOD GETSTARTPOS : LREAL
VAR_INPUT
	LRSETVELOCITY : LREAL;
	LRCLOSEDISTANCE : LREAL;
	LRSETPOSITION : LREAL;
	LRACTPOSITION : LREAL;
	LRCYCLELENGTH : LREAL;
END_VAR
END_METHOD

METHOD HLPDISENGAGECCW
END_METHOD

METHOD HLPDISENGAGECW
END_METHOD

METHOD HLPENGAGECCW
END_METHOD

METHOD HLPENGAGECW
END_METHOD

METHOD INDICATOR
VAR_INPUT
	LRDIFF : LREAL;
	PIINDICATOR : POINTER TO INT;
END_VAR
END_METHOD

METHOD SYNCHRONIZE : LREAL
VAR_INPUT
	LRDIFF : LREAL;
	LRRELPOS : LREAL;
END_VAR
END_METHOD

(* ---- L_MC2P_CLUTCHVELOCITY.fb ---- *)
FUNCTION_BLOCK L_MC2P_CLUTCHVELOCITY
VAR_INPUT
	XENABLE : BOOL;
	XCLOSE : BOOL;
	XOPENINSTANT : BOOL;
	LRCYCVEL : LREAL;
	LRGROUNDVEL : LREAL;
	LRACCDECOPEN : LREAL;
	LRACCDECCLOSE : LREAL;
	LRDECSTOP : LREAL;
	LRJERK : LREAL;
END_VAR
VAR_OUTPUT
	XOPEN : BOOL;
	XCLOSED : BOOL;
	XACCDEC : BOOL;
	LRSETVELOUT : LREAL;
END_VAR
VAR
	HLP_CLUTCHV : L_MC1P_HlpRampGenerator;
	LRBASESPEED : LREAL;
	LRCLOSESPEED : LREAL;
	LRNUMERATOR : LREAL;
	LRDENUMERATOR : LREAL;
	XINITFLAG : BOOL;
	XSETSTARTVELOUT_INT : BOOL;
	XSETSTARTVELOUT_OLD : BOOL;
	LRSTARTVELOUT_INT : LREAL;
	WSTEPCOUNTER : WORD;
	LRSETVELRAMPGENERATOR : LREAL;
	LRLOADRAMPGENDIFF : LREAL;
	XCOMPENSATEVELOCITYJUMP : BOOL;
	XCOMPENSATIONACTIVE : BOOL;
	XLOADCLUTCH_INT : BOOL;
	CLUTCHV_INIT : WORD := 0;
	CLUTCHV_ENABLE : WORD := 1;
	CLUTCHV_CLOSE : WORD := 2;
	CLUTCHV_CLOSING : WORD := 3;
	CLUTCHV_CLOSE_DONE : WORD := 4;
	CLUTCHV_OPENING : WORD := 5;
	CLUTCHV_OPEN_STOP : WORD := 6;
	CLUTCHV_OPENINSTANT_DONE : WORD := 7;
	CLUTCHV_OPENINSTANT_DISABLE : WORD := 8;
	CLUTCHV_CLOSING_STOP : WORD := 9;
	LRSTARTVELOUT : LREAL;
	XSETSTARTVELOUT : BOOL;
END_VAR
END_FUNCTION_BLOCK

METHOD CLUTCHCLOSINGTRANSITION
END_METHOD

METHOD CLUTCHOPENINGTRANSITION
END_METHOD

METHOD COMPENSATEVELOCITYJUMP
END_METHOD

METHOD LOADCLUTCH : BOOL
VAR_INPUT
	XLOADCLUTCH : BOOL;
END_VAR
END_METHOD

METHOD OPENINSTANTTRANSITION
END_METHOD

(* ---- L_MC2P_CONVAXISV.fb ---- *)
FUNCTION_BLOCK L_MC2P_CONVAXISV
VAR_INPUT
	XENABLE : BOOL;
	LRCYCVEL : LREAL;
	DWMODE : DWORD;
	LRCOUPLINGX : LREAL := 1.0;
	LRCOUPLINGY : LREAL := 1.0;
	ETRAVERSINGRANGEX : L_MC1P_TraversingRange;
	ETRAVERSINGRANGEY : L_MC1P_TraversingRange;
	LRCYCLELENGTHY : LREAL;
	LRCYCLELENGTHX : LREAL;
END_VAR
VAR_OUTPUT
	LRSETVELOUT : LREAL;
	XERROR : BOOL;
	EERRORID : L_IE1P_Error;
END_VAR
VAR
	LRSPEED : LREAL := 0;
	LRINPUT : LREAL;
	LRNUM1 : LREAL;
	LRDEN1 : LREAL;
	LRNUM2 : LREAL;
	LRDEN2 : LREAL;
END_VAR
END_FUNCTION_BLOCK

(* ---- L_MC2P_DIFFERENTIATE.fb ---- *)
FUNCTION_BLOCK L_MC2P_DIFFERENTIATE
VAR_INPUT
	LRCYCPOS : LREAL;
	LRCYCLELENGTH : LREAL;
END_VAR
VAR_OUTPUT
	LRSETVELOUT : LREAL;
END_VAR
VAR
	LRPOS : LREAL;
	LRPOSDIFF : LREAL;
	LRLENGTH : LREAL;
	LRPOSOLD : LREAL;
	LRTASKCYCLE : LREAL;
END_VAR
END_FUNCTION_BLOCK

(* ---- L_MC2P_FLEXCAMBASE.fb ---- *)
FUNCTION_BLOCK L_MC2P_FLEXCAMBASE EXTENDS L_MC2P_CamExtendedState
VAR_INPUT
	LRPROFGENMASTERVEL : LREAL;
	LRPROFGENMASTERACC : LREAL;
	LRPROFGENMASTERDEC : LREAL;
	LRPROFGENMASTERJERK : LREAL;
	LRPROFGENSLAVEVEL : LREAL;
	LRPROFGENSLAVEACC : LREAL;
	LRPROFGENSLAVEDEC : LREAL;
	LRPROFGENSLAVEJERK : LREAL;
END_VAR
VAR_OUTPUT
	LRSETOFFSETMASTEROUT : LREAL := 0.0;
	LRSETOFFSETSLAVEOUT : LREAL := 0.0;
END_VAR
VAR
	SCPARPROFILGEN_MASTER : L_MC1P_ProfileParameter;
	SCPARPROFILGEN_SLAVE : L_MC1P_ProfileParameter;
	PROFGEN_MASTER : L_MC1P_PosProfiler;
	PROFGEN_SLAVE : L_MC1P_PosProfiler;
	XPROFGENMASTERCRITICALCYCLE : BOOL;
	XPROFGENMASTERACTIVE : BOOL;
	XPROFGENSALVECRITICALCYCLE : BOOL;
	XPROFGENSLAVEACTIVE : BOOL;
	XEXECUTEPROFGENMASTER : BOOL;
	XEXECUTEPROFGENSLAVE : BOOL;
END_VAR
END_FUNCTION_BLOCK

METHOD CALL_ERRORHANDLER
END_METHOD

METHOD CALL_OUTPUT
END_METHOD

METHOD CALL_PARAMPROFGENMASTER
END_METHOD

METHOD CALL_PARAMPROFGENSLAVE
END_METHOD

METHOD CALL_PROFGENMASTER
END_METHOD

METHOD CALL_PROFGENMASTER_EXECUTECONTROL
END_METHOD

METHOD CALL_PROFGENMASTER_FB
END_METHOD

METHOD CALL_PROFGENMASTER_INPUTOFFSET
END_METHOD

METHOD CALL_PROFGENMASTER_INPUTSCALING
END_METHOD

METHOD CALL_PROFGENMASTER_OUTPUT
END_METHOD

METHOD CALL_PROFGENMASTER_OUTPUTDONE
END_METHOD

METHOD CALL_PROFGENSLAVE
END_METHOD

METHOD CALL_PROFGENSLAVE_EXECUTECONTROL
END_METHOD

METHOD CALL_PROFGENSLAVE_FB
END_METHOD

METHOD CALL_PROFGENSLAVE_INPUTOFFSET
END_METHOD

METHOD CALL_PROFGENSLAVE_INPUTSCALING
END_METHOD

METHOD CALL_PROFGENSLAVE_OUTPUT
END_METHOD

METHOD CALL_RESETOUTPUT
END_METHOD

METHOD CALL_RESETPROFGEN
END_METHOD

METHOD CALL_RESETPROFGENMASTER
END_METHOD

METHOD CALL_RESETPROFGENSLAVE
END_METHOD

METHOD GET_LRPGMASTERSETACCOUT : LREAL
END_METHOD

METHOD GET_LRPGMASTERSETPOSOUT : LREAL
END_METHOD

METHOD GET_LRPGMASTERSETVELOUT : LREAL
END_METHOD

METHOD GET_LRPGSLAVESETACCOUT : LREAL
END_METHOD

METHOD GET_LRPGSLAVESETPOSOUT : LREAL
END_METHOD

METHOD GET_LRPGSLAVESETVELOUT : LREAL
END_METHOD

METHOD GET_XCRITICALCYCLE : BOOL
END_METHOD

METHOD SET_SCALINGINITVAL
END_METHOD

(* ---- L_MC2P_FLEXCAMHIGH.fb ---- *)
FUNCTION_BLOCK L_MC2P_FLEXCAMHIGH EXTENDS L_MC2P_FlexCamState
VAR_INPUT
	XSYNCPOS : BOOL;
	LRSETXPOS : LREAL;
	XHOLDPROFGENMASTER : BOOL;
	XTRIMMASTERPOS : BOOL;
	XTRIMMASTERNEG : BOOL;
	LRPRECTRLGAIN : LREAL := 0;
	LRPRECTRLRATETIME : LREAL := 0;
END_VAR
VAR_OUTPUT
	XSYNCPOSACTIVE : BOOL;
	XENDOFCYCLE : BOOL;
	LRSETMASTERTRIMOFFSETOUT : LREAL := 0.0;
	XPRECTRLACTIVE : BOOL;
	LRPRECTRLACCOUT : LREAL;
END_VAR
VAR
	XSETSTARTXPOS : BOOL;
	LRSETSTARTXPOS : LREAL;
	LRSETMASTERPERIOD : LREAL := 0;
	XSYNCPOS_OLD : BOOL;
	XTRIMMASTERPOS_OLD : BOOL;
	XTRIMMASTERNEG_OLD : BOOL;
	XTRIMMASTERACTIVE : BOOL;
	LRPROFGENMASTERTRIMSTARTPOS : LREAL;
	LROFFSETTRIM_INT : LREAL := 0.0;
	SCCAMTABLE_TMP : MC_Cam_REF;
	SCCAMINFO_TMP : L_MC2P_CamInfo;
	SCPRECTRLSETXPROFILE : L_MC2P_AxisProfile;
	SCPRECTRLSETYPROFILEOUT : L_MC2P_AxisProfile;
	FB_CAMPROFILERRATETIME : L_MC2P_CamBasic;
	XFB_CAMPROFILERRATETIME_PERIODIC : BOOL;
	XFB_CAMPROFILERRATETIME_ERRORCAM : BOOL;
	XFB_CAMPROFILERRATETIME_ERRORIDCAM : L_IE1P_Error;
END_VAR
END_FUNCTION_BLOCK

METHOD CALL_ACCPRECONTROL
END_METHOD

METHOD CALL_ACCPRECONTROL_RATEDACC
END_METHOD

METHOD CALL_CYCLIC_SYNCXTOMASTERPOS
END_METHOD

METHOD CALL_FBMETHODS
END_METHOD

METHOD CALL_OUTPUT
END_METHOD

METHOD CALL_OUTPUT_SETMASTEROFFSETOUT
END_METHOD

METHOD CALL_PARAMPROFGENMASTERTRIMMING
END_METHOD

METHOD CALL_PROFGENMASTER
END_METHOD

METHOD CALL_PROFGENMASTER_INPUTOFFSET
END_METHOD

METHOD CALL_PROFGENMASTER_INPUTSCALING
END_METHOD

METHOD CALL_PROFGENMASTER_INPUTTRIMMING
END_METHOD

METHOD CALL_PROFGENMASTER_OUTPUTDONE
END_METHOD

METHOD CALL_RESETAXISCONVERTER
END_METHOD

METHOD CALL_RESETCOMMANDS
END_METHOD

METHOD CALL_RESETOUTPUT
END_METHOD

METHOD CALL_RESETPROFGEN
END_METHOD

METHOD CALL_SETMASTEROFFSET
END_METHOD

METHOD _CALL_EMPTY
END_METHOD

METHOD CALC_RESTARTXAXIS
END_METHOD

METHOD CALC_XAXIS
END_METHOD

METHOD CALL_OUTPUT_ENDOFPROFILE
END_METHOD

METHOD COPYCAMTABLEID
END_METHOD

METHOD GET_SCCHARCLUTCH : ARRAY [0..1] OF L_MC2P_Characteristics
END_METHOD

METHOD GET_SCPRECTRLSETXPROFILE : L_MC2P_AxisProfile
END_METHOD

METHOD GET_SCPRECTRLSETYPROFILEOUT : L_MC2P_AxisProfile
END_METHOD

METHOD GET_XPGMASTERACTIVE : BOOL
END_METHOD

METHOD SET_MASTERPERIOD
VAR_INPUT
	LRIN : LREAL;
END_VAR
END_METHOD

METHOD SET_STARTXPOS
VAR_INPUT
	LRIN : LREAL;
END_VAR
END_METHOD

METHOD CALL_S000_CYCLIC
END_METHOD

METHOD CALL_S010_01_READY_ENTRY_STATE
END_METHOD

(* ---- L_MC2P_FLEXCAMSTATE.fb ---- *)
FUNCTION_BLOCK L_MC2P_FLEXCAMSTATE EXTENDS L_MC2P_FlexCamBase
VAR_INPUT
	EPOSCTRLDIRECTION : L_MC2P_ReverseCtrlDirection;
END_VAR
VAR
	XDIRECTIONMASTERNEG : BOOL := FALSE;
	XMASTERNOREVERSE : BOOL := FALSE;
	XCLUTCHREVERSE : BOOL;
	XLIMITEDPROFGENMASTER : BOOL;
	LRPROFGENMASTACCDECTIMEDIST : LREAL;
	WCOUNTEREXECUTEPROFGENMASTER : WORD;
	LRMAXVELFREEZE : LREAL;
END_VAR
END_FUNCTION_BLOCK

METHOD CALL_CLUTCHCLOSEMODE
END_METHOD

METHOD CALL_CLUTCHOPENMODE
END_METHOD

METHOD CALL_DETECTDIRECTIONOFMASTER
END_METHOD

METHOD CALL_ERRORHANDLER
END_METHOD

METHOD CALL_OUTPUT
END_METHOD

METHOD CALL_PARAMPROFGENMASTER
END_METHOD

METHOD CALL_PARAMPROFGENMASTERNOREVERSE
END_METHOD

METHOD CALL_PROFGENMASTER
END_METHOD

METHOD CALL_PROFGENMASTERNOTREVERSE
END_METHOD

METHOD CALL_PROFGENMASTER_EXECUTECONTROL
END_METHOD

METHOD CALL_PROFGENMASTER_OUTPUTDONE
END_METHOD

METHOD CALL_PROFGENMASTER_RESTARAFTERSTOP
END_METHOD

METHOD CALL_PROFGENMASTER_STOP
END_METHOD

METHOD CALL_RESETOUTPUT
END_METHOD

METHOD GET_XMASTERPROGENSTOPING : BOOL
END_METHOD

METHOD CALL_PARAMPROFGENMASTERNOTREVERSE
END_METHOD

(* ---- L_MC2P_GEARBOXPOSITION.fb ---- *)
FUNCTION_BLOCK L_MC2P_GEARBOXPOSITION EXTENDS L_MC2P_GearboxPositionBase
VAR_INPUT
	LRCYCLELENGTHX : LREAL;
	LRCYCLELENGTHY : LREAL;
END_VAR
END_FUNCTION_BLOCK

(* ---- L_MC2P_GEARBOXPOSITIONBASE.fb ---- *)
FUNCTION_BLOCK L_MC2P_GEARBOXPOSITIONBASE
VAR_INPUT
	XENABLE : BOOL;
	LRPOSX : LREAL;
	DWNUMERATOR : DWORD := 1;
	DWDENOMINATOR : DWORD := 1;
	XLOADPOSY : BOOL;
	LRLOADPOSY : LREAL;
	LNLOADPOSYRESIDUAL : LINT;
END_VAR
VAR_OUTPUT
	LRPOSY : LREAL;
	LNACTPOSYRESIDUAL : LINT;
	XERROR : BOOL := FALSE;
	EERRORID : L_IE1P_Error := 0;
END_VAR
VAR
	XINIT : BOOL := FALSE;
	LNPOSX : LINT := 0;
	LNPOSY : LINT := 0;
	LNPOSXOLD : LINT := 0;
	LNPOSXDIFF : LINT := 0;
	LNPOSYDIFF : LINT := 0;
	LNPOSYOLD : LINT := 0;
	LNRES_GEARBOX : LINT := 0;
	LRLENX : LREAL;
	LRLENY : LREAL;
	LRLENXOLD : LREAL;
	LRLENYOLD : LREAL;
END_VAR
END_FUNCTION_BLOCK

METHOD CALL_S000_CYCLIC
END_METHOD

METHOD CALL_ERRORHANDLER
END_METHOD

METHOD CALL_RESET
END_METHOD

METHOD L_HLPMODULOADD : LREAL
VAR_INPUT
	LRINPUT : LINT;
	LROFFSET : LINT;
	LRLENGHT : LINT;
END_VAR
END_METHOD

METHOD L_HLPMODULODIFF : LREAL
VAR_INPUT
	LRDIFF : LINT;
	LRLEN : LINT;
END_VAR
END_METHOD

METHOD L_HLPMULDIV : LREAL
VAR_INPUT
	LNINPUT : LINT;
	DWNUMERATOR : DWORD;
	DWDENOMINATOR : DWORD;
	PLNRES : POINTER TO LINT;
END_VAR
END_METHOD

(* ---- L_MC2P_LINEARCOUPLING.fb ---- *)
FUNCTION_BLOCK L_MC2P_LINEARCOUPLING
VAR_INPUT
	XENABLE : BOOL;
	XXRESET : BOOL;
	LRCYCPOSX : LREAL;
	LRSETOFFSETX : LREAL;
	LRCYCLELENGTHX : LREAL;
	LRCYCLELENGTHY : LREAL;
END_VAR
VAR_OUTPUT
	LRSETPOSOUTY : LREAL;
	LRSETVELOUTY : LREAL;
	LRSETVELOUTX : LREAL;
	LRACTPOSX : LREAL;
	XZEROPOS : BOOL;
	XERROR : BOOL;
	EERRORID : L_IE1P_Error;
END_VAR
VAR
	LRPOSDIFF : LREAL;
	LRPOSINPUT : LREAL;
	LRPOSOUTPUT : LREAL;
	LRXLENGTHINT : LREAL;
	LRXLENGTHREST : LREAL;
	XDATAOK : BOOL;
	LRACTXLENGTH : LREAL;
	LRXOFFSETBASE : LREAL;
	LRACTYLENGTH : LREAL;
	XRELOADFLAG : BOOL;
	XENABLEOLD : BOOL;
	LRYSETPOS : INT;
END_VAR
END_FUNCTION_BLOCK

(* ---- L_MC2P_MASTERSLAVESYNC.fb ---- *)
FUNCTION_BLOCK L_MC2P_MASTERSLAVESYNC EXTENDS L_MC2P_Template2Axes_Licence
VAR
	XEXECUTE_INT : BOOL;
	XCONTINUOUSUPDATE_INT : BOOL;
	EBUFFERMODE_INT : MC_BUFFER_MODE := MC_Buffer_Mode.mcAborting;
	XINSYNC_INT : BOOL;
	XBUSY_INT : BOOL;
	XACTIVE_INT : BOOL;
	XCOMMANDABORTED_INT : BOOL;
	XERROR_INT : BOOL;
	EERRORID_INT : L_IE1P_Error;
	ETYPEFUNCTION : L_MC1P_TypeFunction;
	XEXECUTEOLD : BOOL;
	XCOMMANDABORTEDOLD : BOOL;
	PXSOURCEBUFDONE : POINTER TO BOOL;
	XSOURCEBUFDONEOLD : BOOL;
	XRESETOUTPUT : BOOL;
	XCLUTCHACTIVE : BOOL;
	XSUPERIMPOSED : BOOL;
	XCONTINUOUSUPDATE : BOOL;
	XUPDATEBLOCKER : BOOL;
	UIUPDATECOUNTER : UINT;
	DWINSTANCE : __XWORD;
	XBUFFERACTIVE : BOOL;
	WFUNID : WORD;
	XPREVBUFFBDONE : BOOL;
	LRMASTERREFOFFSET : LREAL;
	DWLASTSTEADYSTATE : DWORD;
END_VAR
END_FUNCTION_BLOCK

METHOD CHECKBUFFERMODE
END_METHOD

METHOD CHECK_CONTINUOUSUPDATE
END_METHOD

METHOD CONSIDERMASTERUNSTEADYEVENT
END_METHOD

METHOD GET_SLAVEVALUES
VAR_IN_OUT
	SLAVE : AXIS_REF;
	SCACTVALUESSLAVE : L_MC2P_AxisProfile;
END_VAR
END_METHOD

METHOD READINPUTS
VAR_INPUT
	XREADALL : BOOL;
END_VAR
VAR_IN_OUT
	AXIS : AXIS_REF;
END_VAR
END_METHOD

METHOD RESET_OUTPUTS
END_METHOD

METHOD RESET_OUTPUTSADD
END_METHOD

METHOD RESET_OUTPUTSBYCOMMANDABORTED
END_METHOD

METHOD RESET_OUTPUTSBYERROR
END_METHOD

METHOD SET_BUFFERMODE
END_METHOD

METHOD SET_SLAVEVALUES
VAR_IN_OUT
	SLAVE : AXIS_REF;
	SCSETVALUESSLAVE : L_MC2P_AxisProfile;
END_VAR
END_METHOD

METHOD STOREMASTERSTEADYSTATE
END_METHOD

METHOD SYNCIN
END_METHOD

METHOD FB_INIT : BOOL
VAR_INPUT
	BINITRETAINS : BOOL;
	BINCOPYCODE : BOOL;
END_VAR
END_METHOD

(* ---- L_MC2P_MODIFYAXIS.fb ---- *)
FUNCTION_BLOCK L_MC2P_MODIFYAXIS
VAR
	XBUSY_INT : BOOL;
	XDONE_INT : BOOL;
	XERROR_INT : BOOL;
	EERRORID_INT : L_IE1P_Error;
	L_MC2P_CAMAXISCONVERTER1 : L_MC2P_CamAxisConverter;
	PG : L_MC1P_PosProfiler;
	SCPARAM : L_MC1P_ProfileParameter;
	XRESETOUTPUT : BOOL;
	XEXECUTEOLD : BOOL;
	LRSETSCALING_INT : LREAL;
	LRSETOFFSET_INT : LREAL;
	SCCORRECTAXIS : L_MC2P_AxisProfile;
END_VAR
END_FUNCTION_BLOCK

METHOD OFFSET
VAR_INPUT
	XEXECUTE : BOOL;
	SCINPUTAXIS : L_MC2P_AxisProfile;
	LRSETOFFSET : LREAL;
	EAXISTYPE : L_MC1P_TraversingRange;
	EOFFSETMODE : L_MC2P_OffsetMode;
	LRCYCLETIME : LREAL;
	LRCYCLELENGTH : LREAL;
	LRMAXVELDIFF : LREAL;
	LRMAXACC : LREAL;
	LRMAXDEC : LREAL;
	LRJERK : LREAL;
END_VAR
VAR_OUTPUT
	SCOUTPUTAXIS : L_MC2P_AxisProfile;
	XBUSY : BOOL;
	XDONE : BOOL;
	XERROR : BOOL;
	EERRORID : L_IE1P_Error;
END_VAR
END_METHOD

METHOD SCALING
VAR_INPUT
	XEXECUTE : BOOL;
	SCINPUTAXIS : L_MC2P_AxisProfile;
	LRINPUTAXISPOSOLD : LREAL;
	LRSETSCALING : LREAL;
	XPOSMODE : BOOL;
	EAXISTYPE : L_MC1P_TraversingRange;
	ESCALINGMODE : L_MC2P_ScalingMode;
	LRCYCLETIME : LREAL;
	LRCYCLELENGTH : LREAL;
	LRMAXVELDIFF : LREAL;
	LRMAXACC : LREAL;
	LRMAXDEC : LREAL;
	LRJERK : LREAL;
END_VAR
VAR_OUTPUT
	SCOUTPUTAXIS : L_MC2P_AxisProfile;
	XBUSY : BOOL;
	XDONE : BOOL;
	XERROR : BOOL;
	EERRORID : L_IE1P_Error;
END_VAR
END_METHOD

METHOD CALC_AXISVALUESWITHOFFSET
VAR_INPUT
	SCINPUTAXIS : L_MC2P_AxisProfile;
	EAXISTYPE : L_MC1P_TraversingRange;
	LRCYCLELENGTH : LREAL;
END_VAR
VAR_OUTPUT
	SCOUTPUTAXIS : L_MC2P_AxisProfile;
END_VAR
END_METHOD

METHOD SET_PROFILEGENERATORWITHOFFSET
VAR_INPUT
	LRCYCLETIME : LREAL;
	LRSETOFFSET : LREAL;
	LRSETOFFSET_INT : LREAL;
	LRMAXVELDIFF : LREAL;
	LRMAXACC : LREAL;
	LRMAXDEC : LREAL;
	LRJERK : LREAL;
END_VAR
END_METHOD

METHOD CALC_AXISVALUESWITHSCALING
VAR_INPUT
	SCINPUTAXIS : L_MC2P_AxisProfile;
	EAXISTYPE : L_MC1P_TraversingRange;
END_VAR
VAR_OUTPUT
	SCOUTPUTAXIS : L_MC2P_AxisProfile;
END_VAR
END_METHOD

METHOD GETSCALEDAXISPOSITION : LREAL
VAR_INPUT
	LRPOS : LREAL;
END_VAR
END_METHOD

METHOD SET_CAMAXISCONVERTERWITHSCALING
VAR_INPUT
	ESCALINGMODE : L_MC2P_ScalingMode;
	EAXISTYPE : L_MC1P_TraversingRange;
	LRCYCLELENGTH : LREAL;
	LRINPUTAXISPOS : LREAL;
	LRINPUTAXISPOSOLD : LREAL;
END_VAR
END_METHOD

METHOD SET_PROFILEGENERATORWITHSCALING
VAR_INPUT
	SCINPUTAXIS : L_MC2P_AxisProfile;
	XPOSMODE : BOOL;
	LRCYCLETIME : LREAL;
	ESCALINGMODE : L_MC2P_ScalingMode;
	LRSCALINGFACTOR : LREAL;
	LRMAXVELDIFF : LREAL;
	LRMAXACC : LREAL;
	LRMAXDEC : LREAL;
	LRJERK : LREAL;
END_VAR
END_METHOD

METHOD CALL_PROFILEGENERATOR
END_METHOD

METHOD RESET_INTERNOFFSETSCALING
END_METHOD

METHOD RESET_OUTPUTS
END_METHOD

METHOD RESET_PROFILEGENERATORVALUES
END_METHOD

METHOD SET_INTERNOFFSET
VAR_INPUT
	LRSETOFFSETPOS_INT : LREAL;
	LRSETOFFSETVEL_INT : LREAL;
	LRSETOFFSETACC_INT : LREAL;
END_VAR
END_METHOD

METHOD SET_OUTPUTS
VAR_OUTPUT
	XBUSY : BOOL;
	XDONE : BOOL;
	XERROR : BOOL;
	EERRORID : L_IE1P_Error;
END_VAR
END_METHOD

(* ---- L_MC2P_MULTICAMSEQUENCER.fb ---- *)
FUNCTION_BLOCK L_MC2P_MULTICAMSEQUENCER
VAR_INPUT
	XENABLE : BOOL;
	XCAMSEQUENCER : BOOL;
	EMODE : L_MC2P_CamSequenceMode;
	XCAMCHANGEINSTANT : BOOL;
	ESETCAMTABLE : L_MC2P_CamTable;
	XENDOFPROFILEIN : BOOL;
	CAMTABLE1 : MC_CAM_REF;
	CAMTABLE2 : MC_CAM_REF;
	CAMTABLE3 : MC_CAM_REF;
	CAMTABLE4 : MC_CAM_REF;
END_VAR
VAR_OUTPUT
	XDONE : BOOL;
	XBUSY : BOOL;
	XERROR : BOOL;
	EERRORID : L_IE1P_Error;
	ESETCAMTABLEOUT : L_MC2P_CamTable;
	CAMTABLEOUT : MC_CAM_REF;
END_VAR
VAR
	EFMSTATE : L_MC2P_States := L_MC2P_States.INIT;
	XINITSTATE : BOOL;
	XENABLE_OLD : BOOL;
	XLOADCAMTABLE_OLD : BOOL;
	XENDOFPROFILEIN_OLD : BOOL;
	XCAMSEQUENCER_OLD : BOOL;
	XCAMCHANGEINSTANT_OLD : BOOL;
	XCAMSEQUENCERACTIVE : BOOL;
END_VAR
END_FUNCTION_BLOCK

METHOD CALL_ERRORHANDLER
END_METHOD

METHOD CALL_FBMETHODS
END_METHOD

METHOD CALL_OUTPUT
END_METHOD

METHOD CALL_RESETCOMMANDS
END_METHOD

METHOD CALL_RESETOUTPUT
END_METHOD

METHOD CALL_STATEMACHINE
END_METHOD

METHOD CALL_SETCAMTABLEOUT
VAR_INPUT
	ESETCAMTABLE : L_MC2P_CamTable;
END_VAR
END_METHOD

METHOD CAMREFCHANGED : BOOL
VAR_IN_OUT
	CAMREFNEW : MC_CAM_REF;
	CAMREFOLD : MC_CAM_REF;
END_VAR
END_METHOD

METHOD CALL_S000_CYCLIC
END_METHOD

METHOD CALL_S001_INIT
END_METHOD

METHOD CALL_S002_READY
END_METHOD

METHOD CALL_S151_SEQUENCE_CYCLICCAM1
END_METHOD

METHOD CALL_S152_SEQUENCE_CYCLICCAM3
END_METHOD

METHOD CALL_S153_SEQUENCE_CAM1CYCLICCAM3CAM1
END_METHOD

METHOD CALL_S154_SEQUENCE_CAM1CAM2CYCLICCAM3CAM4CAM1
END_METHOD

(* ---- L_MC2P_PHASING.fb ---- *)
FUNCTION_BLOCK L_MC2P_PHASING EXTENDS L_MC2P_Template2Axes_Licence
VAR_INPUT
	EXECUTE : BOOL;
	PHASESHIFT : LREAL := 0;
	VELOCITY : LREAL := 3600.0;
	ACCELERATION : LREAL := 3600.0;
	DECELERATION : LREAL := 3600.0;
	JERK : LREAL := 0.0;
	BUFFERMODE : MC_BUFFER_MODE := MC_Buffer_Mode.mcAborting;
END_VAR
VAR_OUTPUT
	DONE : BOOL;
	BUSY : BOOL;
	ACTIVE : BOOL;
	COMMANDABORTED : BOOL;
	ERROR : BOOL;
	ERRORID : L_IE1P_Error;
END_VAR
VAR
	L_MC2P_MODIFYAXIS1 : L_MC2P_ModifyAxis;
	XSUPERIMPOSED : BOOL;
	WFUNID : WORD;
	SCINPUTMASTERSOURCE : L_MC2P_AxisProfile;
	SCOUTPUTSLAVE : L_MC2P_AxisProfile;
	XEXECUTEOLD : BOOL;
	XRESETOUTPUT : BOOL;
	DWINSTANCE : __XWORD;
	XBUFFERACTIVE : BOOL;
	XPREVBUFFBDONE : BOOL;
	LRPHASESHIFT_INT : LREAL;
	LRVELOCITY_INT : LREAL;
	LRACCELERATION_INT : LREAL;
	LRDECELERATION_INT : LREAL;
	LRJERK_INT : LREAL;
	EBUFFERMODE_INT : MC_BUFFER_MODE;
	XRELATIVE : BOOL;
	ETYPEFUNCTION : L_MC1P_TypeFunction;
	LRACTPHASESHIFT : LREAL;
	LRPHASESHIFTOLD : LREAL;
	LRPHASESHIFTSET : LREAL;
	XCOMMANDABORTEDOLD : BOOL;
	PXDUMMY : POINTER TO BOOL;
END_VAR
END_FUNCTION_BLOCK

METHOD GET_MASTERVALUES
END_METHOD

METHOD INIT_PHASING
END_METHOD

METHOD READINPUTS
VAR_INPUT
	XREADALL : BOOL;
END_VAR
VAR_IN_OUT
	AXIS : AXIS_REF;
END_VAR
END_METHOD

METHOD RESET_OUTPUTS
END_METHOD

METHOD RESET_OUTPUTSBYCOMMANDABORTED
END_METHOD

METHOD RESET_OUTPUTSBYERROR
END_METHOD

METHOD SET_BUFFERMODE
END_METHOD

(* ---- L_MC2P_READLMDFILE.fb ---- *)
FUNCTION_BLOCK L_MC2P_READLMDFILE
VAR_OUTPUT
	XNEWDATAAVAILABLE : BOOL;
END_VAR
VAR
	SFILE_INT : STRING := '';
	EDATA_INT : L_MC2P_LMData;
	PDATA_INT : POINTER TO BYTE;
	WDATAELEMENTS_INT : WORD;
	XENABLEONLINECHANGE_INT : BOOL;
	XBUSY_INT : BOOL;
	XDONE_INT : BOOL;
	XERROR_INT : BOOL;
	EERRORID_INT : L_IE1P_Error;
	XEXECUTEOLD : BOOL;
	HFILE : SYSFILE.RTS_IEC_HANDLE;
	RES : SYSFILE.RTS_IEC_RESULT;
	ID : L_MC2P_Magic;
	DWLENGTH : DWORD;
	XACTIVECRYPTING : BOOL;
	CRYPT : Crypting;
	CK : ARRAY [0..3] OF ULINT;
	CCYCLES : WORD;
	DIRAWDATAREAD : DINT;
	DWSTARTCDATA : DWORD;
	ABDATA : ARRAY [0..15] OF BYTE;
	DATAIDX : DWORD;
	AVAILABLEDATA : DWORD;
	XDATAREADDONE : BOOL;
	UDIFSIZE : UDINT;
	UDIFBYTESREAD : UDINT;
	ITFCALLBACK : CmpEventMgr.ICmpEventCallback;
	HEVENTDOWNLOADDONE : SysTypes.RTS_IEC_HANDLE;
	HINTERFACEDOWNLOADDONE : SysTypes.RTS_IEC_HANDLE;
	HEVENTBOOTPROJECTLOADED : SysTypes.RTS_IEC_HANDLE;
	HINTERFACEBOOTPROJECTLOADED : SysTypes.RTS_IEC_HANDLE;
	HEVENTRESETDONE : SysTypes.RTS_IEC_HANDLE;
	HINTERFACERESETDONE : SysTypes.RTS_IEC_HANDLE;
	HEVENTDOWNLOADSINGLEFILE : SysTypes.RTS_IEC_HANDLE;
	HINTERFACEDOWNLOADSINGLEFILE : SysTypes.RTS_IEC_HANDLE;
	DWEVENTCOUNTER : DWORD;
	XDATAVALID : BOOL;
	XDATAACTIVE : BOOL;
	DWDATACRC : DWORD;
	LRACTXPOS : LREAL;
	XDUMMY : BOOL;
END_VAR
END_FUNCTION_BLOCK

METHOD CHECKFILENAME : BOOL
VAR_IN_OUT
	SFILE : STRING;
END_VAR
END_METHOD

METHOD CHECKINPUTS : BOOL
END_METHOD

METHOD LOADDATA
END_METHOD

METHOD MAIN
END_METHOD

METHOD READFRAMES
VAR_INPUT
	HFILE : SYSFILE.RTS_IEC_HANDLE;
END_VAR
END_METHOD

METHOD READORGA
VAR_INPUT
	HFILE : SYSFILE.RTS_IEC_HANDLE;
END_VAR
END_METHOD

METHOD READSPECIFICDATA
VAR_INPUT
	HFILE : SYSFILE.RTS_IEC_HANDLE;
END_VAR
END_METHOD

METHOD RESET
END_METHOD

METHOD CHECKCRC : BOOL
VAR_INPUT
	HFILE : SYSFILE.RTS_IEC_HANDLE;
	DWLENGTH : DWORD;
END_VAR
END_METHOD

METHOD CRCCHECKSUM32BITINCREMENTAL : DWORD
VAR_INPUT
	PBDATA : POINTER TO BYTE;
	DWDATASIZE : DWORD;
	DWCRC : DWORD;
END_VAR
END_METHOD

METHOD EVENTCALLBACK : UDINT
VAR_INPUT
	PEVENTPARAM : POINTER TO EventParam;
END_VAR
END_METHOD

METHOD REGISTEREVENT
END_METHOD

METHOD UNREGISTEREVENT
END_METHOD

METHOD RESETREADDATA
END_METHOD

METHOD CREADCHAR : STRING(16)
VAR_INPUT
	HFILE : SYSFILE.RTS_IEC_HANDLE;
	N : UINT;
END_VAR
END_METHOD

METHOD CREADF64 : LREAL
VAR_INPUT
	HFILE : SYSFILE.RTS_IEC_HANDLE;
END_VAR
END_METHOD

METHOD CREADU16 : WORD
VAR_INPUT
	HFILE : SYSFILE.RTS_IEC_HANDLE;
END_VAR
END_METHOD

METHOD CREADU32 : DWORD
VAR_INPUT
	HFILE : SYSFILE.RTS_IEC_HANDLE;
END_VAR
END_METHOD

METHOD READCRYPTDATA : DWORD
VAR_INPUT
	HFILE : SYSFILE.RTS_IEC_HANDLE;
	DWSIZE : DWORD;
END_VAR
VAR_IN_OUT
	DATA : L_MC2P_IntData;
END_VAR
END_METHOD

METHOD GETNEXTFRAME
VAR_INPUT
	HFILE : SYSFILE.RTS_IEC_HANDLE;
	DWOFFSET : DWORD;
END_VAR
END_METHOD

METHOD READ
VAR_INPUT
	HFILE : SYSFILE.RTS_IEC_HANDLE;
	PBYBUFFER : POINTER TO BYTE;
	ULSIZE : UINT;
END_VAR
VAR_OUTPUT
	UDIDATAREAD : UDINT;
END_VAR
END_METHOD

METHOD READCHAR : STRING(16)
VAR_INPUT
	HFILE : SYSFILE.RTS_IEC_HANDLE;
	N : UINT;
END_VAR
END_METHOD

METHOD READF64 : LREAL
VAR_INPUT
	HFILE : SYSFILE.RTS_IEC_HANDLE;
END_VAR
END_METHOD

METHOD READU16 : WORD
VAR_INPUT
	HFILE : SYSFILE.RTS_IEC_HANDLE;
END_VAR
END_METHOD

METHOD READU32 : DWORD
VAR_INPUT
	HFILE : SYSFILE.RTS_IEC_HANDLE;
END_VAR
END_METHOD

METHOD FB_EXIT : BOOL
VAR_INPUT
	BINCOPYCODE : BOOL;
END_VAR
END_METHOD

METHOD FB_INIT : BOOL
VAR_INPUT
	BINITRETAINS : BOOL;
	BINCOPYCODE : BOOL;
END_VAR
END_METHOD

METHOD ABORT : UDINT
END_METHOD

METHOD EXECUTE : UDINT
END_METHOD

(* ---- L_MC2P_RESETPHASING.fb ---- *)
FUNCTION_BLOCK L_MC2P_RESETPHASING EXTENDS L_MC2P_TemplateAxis_Licence
VAR_INPUT
	XEXECUTE : BOOL;
END_VAR
VAR_OUTPUT
	XDONE : BOOL;
	XERROR : BOOL;
	EERRORID : L_IE1P_Error;
END_VAR
VAR
	XEXECUTEOLD : BOOL;
	PXDUMMY : POINTER TO BOOL;
END_VAR
END_FUNCTION_BLOCK

(* ---- L_MC2P_TAPPETDATAOBJECT.fb ---- *)
FUNCTION_BLOCK L_MC2P_TAPPETDATAOBJECT
VAR_INPUT
	DWSTRUCTID : DWORD := L_MC2P_Constants.gC_dwCheckIDTappet;
	LRTAPPETON : LREAL;
	LRTAPPETOFF : LREAL;
END_VAR
VAR
	BASE : POINTER TO BYTE;
	DATATYPE : L_MC2P_MotionDataType;
	SIZE : UDINT;
	STARTADRESS : POINTER TO BYTE;
END_VAR
END_FUNCTION_BLOCK

(* ---- L_MC2P_TAPPETDATAPOS.fb ---- *)
FUNCTION_BLOCK L_MC2P_TAPPETDATAPOS
VAR_INPUT
	DWSTRUCTID : DWORD := L_MC2P_Constants.gC_dwCheckIDTappetPos;
	LRTAPPETON : LREAL;
	LRTAPPETOFF : LREAL;
END_VAR
VAR
	BASE : POINTER TO BYTE;
	DATATYPE : L_MC2P_MotionDataType;
	SIZE : UDINT;
	STARTADRESS : POINTER TO BYTE;
END_VAR
END_FUNCTION_BLOCK

(* ---- L_MC2P_TAPPETDATATIME.fb ---- *)
FUNCTION_BLOCK L_MC2P_TAPPETDATATIME
VAR_INPUT
	DWSTRUCTID : DWORD := L_MC2P_Constants.gC_dwCheckIDTappetTime;
	LRTAPPETON : LREAL;
	LRTAPPETTIME : LREAL;
END_VAR
VAR
	BASE : POINTER TO BYTE;
	DATATYPE : L_MC2P_MotionDataType;
	SIZE : UDINT;
	STARTADRESS : POINTER TO BYTE;
END_VAR
END_FUNCTION_BLOCK

(* ---- L_MC2P_TAPPETREFFROMFILE.fb ---- *)
FUNCTION_BLOCK L_MC2P_TAPPETREFFROMFILE EXTENDS L_MC2P_ReadLMDFile
VAR_INPUT
	XEXECUTE : BOOL;
	SFILENAME : STRING := '';
	ITFTAPPETDATA : L_MC2P_ITappetData;
	UDITAPPETDATACOUNT : UDINT;
	XRELOADABLE : BOOL;
END_VAR
VAR_OUTPUT
	XDONE : BOOL;
	XBUSY : BOOL;
	XERROR : BOOL;
	EERRORID : L_IE1P_Error;
END_VAR
VAR
	MOTIONDATA_INT : L_MC2P_ITappetData;
	SCTAPPETDATA : L_MC2P_TappetData;
	XRELOADOLD : BOOL;
	RELOAD : BOOL;
END_VAR
END_FUNCTION_BLOCK

METHOD CHECKFILENAME : BOOL
VAR_IN_OUT
	SFILE : STRING;
END_VAR
END_METHOD

METHOD CHECKINPUTS : BOOL
END_METHOD

METHOD LOADDATA
END_METHOD

METHOD MAIN
END_METHOD

METHOD GETID : DWORD
END_METHOD

METHOD GETTAPPETDATA : POINTER TO L_MC2P_TappetData
END_METHOD

METHOD SETCAMDATAACTIVE
VAR_INPUT
	XCAMACITVE : BOOL;
END_VAR
END_METHOD

METHOD SETMASTERVALUES
VAR_INPUT
	LRMASTERPOS : LREAL;
END_VAR
END_METHOD

METHOD GETTAPPET
VAR_INPUT
	HFILE : SYSFILE.RTS_IEC_HANDLE;
	ITFCAMDATA : L_MC2P_ITappetData;
	WDATAELEMENTS : WORD;
	DWCOUNT : DWORD;
END_VAR
END_METHOD

METHOD READSPECIFICDATA
VAR_INPUT
	HFILE : SYSFILE.RTS_IEC_HANDLE;
END_VAR
END_METHOD

METHOD READTAPPETDATA
VAR_INPUT
	HFILE : SYSFILE.RTS_IEC_HANDLE;
END_VAR
END_METHOD

(* ---- L_MC2P_TAPPETREFFROMSTRUCT.fb ---- *)
FUNCTION_BLOCK L_MC2P_TAPPETREFFROMSTRUCT EXTENDS L_MC2P_TemplateNoAxis
VAR_INPUT
	XEXECUTE : BOOL;
	SNAME : STRING(50);
	ETAPPETTYPE : L_MC2P_TappetType;
	UDICAMDATACOUNT : UDINT;
	LRXSTARTPOS : LREAL;
	LRXENDPOS : LREAL;
	ITFTAPPETDATA : L_MC2P_ITappetData;
END_VAR
VAR_OUTPUT
	XDONE : BOOL;
	XBUSY : BOOL;
	XERROR : BOOL;
	EERRORID : L_IE1P_Error;
END_VAR
VAR
	I : UDINT;
	SCDATA : L_MC2P_TappetData;
	PDATAPOS : POINTER TO L_MC2P_TappetDataPos;
	PDATATIME : POINTER TO L_MC2P_TappetDataTime;
	DWGUID : DWORD;
	XEXECUTEOLD : BOOL;
	XRESETOUTPUT : BOOL;
	XDATAVALID : BOOL;
	XDATAACTIVE : BOOL;
	DWDATACRC : DWORD;
	LRACTXPOS : LREAL;
END_VAR
END_FUNCTION_BLOCK

METHOD GETID : DWORD
END_METHOD

METHOD GETTAPPETDATA : POINTER TO L_MC2P_TappetData
END_METHOD

METHOD SETCAMDATAACTIVE
VAR_INPUT
	XCAMACITVE : BOOL;
END_VAR
END_METHOD

METHOD SETMASTERVALUES
VAR_INPUT
	LRMASTERPOS : LREAL;
END_VAR
END_METHOD

(* ---- L_MC2P_TAPPETREFTOFILE.fb ---- *)
FUNCTION_BLOCK L_MC2P_TAPPETREFTOFILE EXTENDS L_MC2P_WriteLMDFile
VAR_INPUT
	XEXECUTE : BOOL;
	SFILENAME : STRING := '';
	ITFTAPPETTABLE : L_MC2P_Tappet_REF;
END_VAR
VAR_OUTPUT
	XDONE : BOOL;
	XBUSY : BOOL;
	XERROR : BOOL;
	EERRORID : L_IE1P_Error;
END_VAR
VAR
	XRELOADOLD : BOOL;
	RELOAD : BOOL;
END_VAR
END_FUNCTION_BLOCK

METHOD MAIN
END_METHOD

METHOD WRITESPECIFICDATA
VAR_INPUT
	HFILE : SYSFILE.RTS_IEC_HANDLE;
END_VAR
END_METHOD

METHOD WRITETAPPET
VAR_INPUT
	HFILE : SYSFILE.RTS_IEC_HANDLE;
	ITFCAMDATA : L_MC2P_ITappetData;
	DWCOUNT : DWORD;
END_VAR
END_METHOD

METHOD WRITETAPPETDATA
VAR_INPUT
	HFILE : SYSFILE.RTS_IEC_HANDLE;
END_VAR
END_METHOD

(* ---- L_MC2P_TAPPETREGISTER.fb ---- *)
FUNCTION_BLOCK L_MC2P_TAPPETREGISTER EXTENDS L_MC2P_TemplateAxis_Licence
VAR_INPUT
	XENABLE : BOOL;
	XFORCE : BOOL;
	ITFTAPPETTABLE : L_MC2P_Tappet_Ref;
	LROFFSET : LREAL;
	LRHYSTERESE : LREAL;
	LRREACTTIMEON : LREAL;
	LRREACTTIMEOFF : LREAL;
	EVALUESOURCE : MC_SOURCE;
	BYDIGITALOUTPUTSEL : BYTE := 0;
	PFASTIO_OUT : POINTER TO L_FastIO_OutRef;
	XOUTPUTSTATE : BOOL := TRUE;
	XEDGECONTROL : BOOL;
END_VAR
VAR_OUTPUT
	XSWITCH : BOOL;
	XBUSY : BOOL;
	XERROR : BOOL;
	EERRORID : L_IE1P_Error;
	BYTAPPETNO : BYTE;
	LRTIMEONRELATIVE : LREAL;
	LRTIMEOFFRELATIVE : LREAL;
END_VAR
VAR
	L_MC1P_ZERODETECT1 : L_MC1P_ZeroDetect;
	PDWABSOLUTECOUNTER : POINTER TO DWORD;
	DWDUMMYCOUNTER : DWORD;
	XMAPPINGINIT : BOOL;
	LRTIMERTICK : LREAL;
	LRTIMERTICKOFF : ARRAY [0..3] OF LREAL;
	LRTIMERPOSOFFSET : ARRAY [0..3] OF LREAL;
	LRFASTIOEXTRA : LREAL := 4.0;
	DWABSOLUTECOUNTEROLD : DWORD;
	DIMAPPINGCOUNT : DINT;
	WTIMERON : WORD;
	WTIMEROFF : WORD;
	XENABLEOLD : BOOL;
	XRESETOUTPUT : BOOL;
	SCDATAOBJECT_INT : ARRAY [0..L_MC2P_InternalConst.C_TAPPETS_BUFFERSIZE] OF L_MC2P_TappetDataObject;
	SCONOFF : ARRAY [0..L_MC2P_InternalConst.C_TAPPETS_BUFFERSIZE] OF L_MC2P_TappetDataObject;
	AXCAMSWITCHEDON : ARRAY [0..L_MC2P_InternalConst.C_TAPPETS_BUFFERSIZE] OF BOOL;
	AICAMSWITCHONCYCLE : ARRAY [0..L_MC2P_InternalConst.C_TAPPETS_BUFFERSIZE] OF INT;
	AXCAMSWITCHEDOFF : ARRAY [0..L_MC2P_InternalConst.C_TAPPETS_BUFFERSIZE] OF BOOL;
	AICAMSWITCHOFFCYCLE : ARRAY [0..L_MC2P_InternalConst.C_TAPPETS_BUFFERSIZE] OF INT;
	ICYCLE : INT;
	ICYCLEFAST : INT;
	PSCTAPPETDATA_INT : POINTER TO L_MC2P_TappetData;
	DWGUID_INT : DWORD;
	LROFFSET_INT : LREAL;
	LRHYTERESE_INT : LREAL;
	LRREACTTIMEON_INT : LREAL;
	LRREACTTIMEOFF_INT : LREAL;
	EVALUESOURCE_INT : MC_SOURCE;
	LRGETPOSITION : LREAL;
	LRGETPOSITIONOLD : LREAL;
	LRCYCLELENGTH : LREAL;
	LRPOSDIFF : LREAL;
	BYDIRECTION : BYTE;
	XOFFSETCHANGE : BOOL;
	LRTAPPETON_INT : ARRAY [0..L_MC2P_InternalConst.C_TAPPETS_BUFFERSIZE] OF LREAL;
	LRTAPPETOFF_INT : ARRAY [0..L_MC2P_InternalConst.C_TAPPETS_BUFFERSIZE] OF LREAL;
	XTAPPETOK : BOOL;
	LRGETPOSITIONOLDINIT : LREAL;
	BYSTEPFASTIO : BYTE;
	BYDIRECTIONSAVE : BYTE;
	XSWITCHFASTIO : BOOL;
	UDIFASTIOORDER : UDINT;
	XFASTIOORDERSTOP : BOOL;
	BYI : BYTE;
	XFORCEFASTAKTIV : BOOL;
	UDIDX1 : UDINT;
	UDISTART1 : UDINT;
	LRINTPOSOLD : LREAL;
	XORDERPAUSE : BOOL;
	BYDIRECTIONOLD : BYTE;
	BYTAPPETIMEAKTIVE : BYTE;
	LRSWITCHTIME : LREAL;
	XTIMERSTART : BOOL;
	UDIFLAGTAPPETNO : UDINT;
	WRINGBUFFERINDEX : WORD;
	LRVELRINGBUFFER : ARRAY [0..wEncFilterCycles] OF LREAL;
	LRVELFILTERBUFFERSUM : LREAL;
	LRPOSDIFFINFILT : LREAL;
	XFLAGBUFFERFULL : BOOL;
	LRPOSDIFFHYST : LREAL;
	XHYSTERESEACTIVE : BOOL;
	XFORCEACTIVE : BOOL;
	PFREEENCODERAXIS : POINTER TO _Axis_Ref_Enc;
	EENCTYPE : L_Mc1P_EncoderType;
	LRDELAYCOMPPLCCYCLES : LREAL := 0.0;
	UDIFORINIT : UDINT;
	LRSWITCHDIFFOLD : LREAL;
	RES : INT;
	XTAPPETFREE : BOOL;
	XTAPPETOKOLD : BOOL;
	XZERO : BOOL;
	XTAPPETCLOSED : BOOL;
	XINITEDGECON : BOOL;
	XSETDELAYCOMP : BOOL;
	DWSTEADYSTATEOLD : DWORD;
	XSETDELAYCOMPOLD : BOOL;
	XDIRECTIONDETECT : BOOL;
	WCOUNTCW : WORD;
	WCOUNTCCW : WORD;
	WCOUNTMAX : WORD := 10;
	EDIRECTIONTMP : L_MC2P_Direction;
	BYDIRECTIONTMP : BYTE;
	WENCFILTERCYCLES : WORD := 10;
	LRFASTIO_OFFSETTIME : LREAL := 3;
	LRVELOCITY : LREAL;
END_VAR
END_FUNCTION_BLOCK

METHOD CALCPOSTPONE : INT
VAR_INPUT
	LRDYNAMIZE : LREAL;
	LRON : LREAL;
	LROFF : LREAL;
	LRLEN : LREAL;
END_VAR
END_METHOD

METHOD CALCTAPPETPOS : BOOL
END_METHOD

METHOD CALCTAPPETTIME : BOOL
END_METHOD

METHOD CHECKINPUTDATA : BOOL
VAR_IN_OUT
	AXIS : AXIS_REF;
END_VAR
END_METHOD

METHOD CHECKINPUTSTRUCT : BOOL
VAR_IN_OUT
	AXIS : AXIS_REF;
END_VAR
END_METHOD

METHOD CLEARMEMINTERN
END_METHOD

METHOD DIRECTIONFORCE
VAR_INPUT
	WAXISSTATE : L_MC1P_AXIS_STATE;
END_VAR
END_METHOD

METHOD DIRECTIONHYST
VAR_IN_OUT
	AXIS : AXIS_REF;
END_VAR
END_METHOD

METHOD DYNAMIZE : LREAL
VAR_INPUT
	REACTTIME : LREAL;
END_VAR
END_METHOD

METHOD GETABSOLUTECOUNTER
END_METHOD

METHOD GETPOSITION : LREAL
VAR_INPUT
	EVALUESOURCE : MC_SOURCE;
END_VAR
END_METHOD

METHOD INSERTENTRYINTOFIFO : INT
VAR_INPUT
	LRTIMERTICK : LREAL;
	BSTATE : BOOL;
END_VAR
END_METHOD

METHOD READINPUTS : BOOL
VAR_IN_OUT
	AXIS : AXIS_REF;
END_VAR
END_METHOD

METHOD RESET
END_METHOD

METHOD RESET_OUTPUTSBYERROR
VAR_INPUT
	XERROR : BOOL;
END_VAR
END_METHOD

METHOD SWITCHFASTIO
VAR_INPUT
	BYDIGITALOUTPUTSEL : BYTE;
	XHYSTERESEACTIVE : BOOL;
	LRDELAYCOM : LREAL;
END_VAR
END_METHOD

METHOD SWITCHTAPPET : BOOL
VAR_INPUT
	XENABLE : BOOL;
END_VAR
END_METHOD

METHOD CHECKDYNAMIZE : BOOL
VAR_INPUT
	LRDYNAMIZE : LREAL;
END_VAR
END_METHOD

METHOD CHECKPOS : LREAL
VAR_INPUT
	LRPOS : LREAL;
END_VAR
END_METHOD

METHOD CHECKTIME : BOOL
VAR_INPUT
	LRDYNAMIZE : LREAL;
END_VAR
END_METHOD

(* ---- L_MC2P_TEMPLATE2AXES.fb ---- *)
FUNCTION_BLOCK L_MC2P_TEMPLATE2AXES
VAR_INPUT
	MASTER : L_MC1P_IAXIS_REF_MASTERVALUES;
END_VAR
VAR_IN_OUT
	SLAVE : AXIS_REF;
END_VAR
VAR
	SINSTANCESTR : STRING;
	XERROROLD : BOOL;
	WERRORIDOLD : WORD;
	DWERRORITFID : DWORD;
	ITFMASTERVALUESDUMMY : L_MC1P_AxisMasterValuesEmpty;
END_VAR
END_FUNCTION_BLOCK

METHOD FB_GETERRORITFID : DWORD
END_METHOD

METHOD FB_RESETERROR
VAR_INPUT
	XERROR : BOOL;
	WERRORID : WORD;
END_VAR
END_METHOD

METHOD FB_SETERROR
VAR_INPUT
	WERRORID : WORD := 0;
	XSETERRORSTOP : BOOL := FALSE;
END_VAR
END_METHOD

METHOD FB_INIT : BOOL
VAR_INPUT
	BINITRETAINS : BOOL;
	BINCOPYCODE : BOOL;
END_VAR
END_METHOD

(* ---- L_MC2P_TEMPLATE2AXES_LICENCE.fb ---- *)
FUNCTION_BLOCK L_MC2P_TEMPLATE2AXES_LICENCE EXTENDS L_MC2P_Template2Axes
VAR
	LICHANDLING : L_IMHP_LLMHandling;
END_VAR
END_FUNCTION_BLOCK

METHOD ACTIVATEAPPCREDIT : BOOL
VAR_INPUT
	XACTIVATE : BOOL;
END_VAR
END_METHOD

(* ---- L_MC2P_TEMPLATE3AXES.fb ---- *)
FUNCTION_BLOCK L_MC2P_TEMPLATE3AXES
VAR_IN_OUT
	MASTER1 : AXIS_REF;
	MASTER2 : AXIS_REF;
	SLAVE : AXIS_REF;
END_VAR
VAR
	SINSTANCESTR : STRING;
	XERROROLD : BOOL;
	WERRORIDOLD : WORD;
	DWERRORITFID : DWORD;
END_VAR
END_FUNCTION_BLOCK

METHOD FB_GETERRORITFID : DWORD
END_METHOD

METHOD FB_RESETERROR
VAR_INPUT
	XERROR : BOOL;
	WERRORID : WORD;
END_VAR
END_METHOD

METHOD FB_SETERROR
VAR_INPUT
	WERRORID : WORD := 0;
	XSETERRORSTOP : BOOL := FALSE;
END_VAR
END_METHOD

METHOD FB_INIT : BOOL
VAR_INPUT
	BINITRETAINS : BOOL;
	BINCOPYCODE : BOOL;
END_VAR
END_METHOD

(* ---- L_MC2P_TEMPLATE3AXES_LICENCE.fb ---- *)
FUNCTION_BLOCK L_MC2P_TEMPLATE3AXES_LICENCE EXTENDS L_MC2P_Template3Axes
VAR
	LICHANDLING : L_IMHP_LLMHandling;
END_VAR
END_FUNCTION_BLOCK

METHOD ACTIVATEAPPCREDIT : BOOL
VAR_INPUT
	XACTIVATE : BOOL;
END_VAR
END_METHOD
